// TIA Portal project "汽车系统" (V15.1)
// 汽车雨刷与车窗系统

(* hardware
DEVICE "S7-1200 station_1"  S7-1200 Station
   slot 0: "Rack_0"  S7-1200 Rack  Rack  V1.0
   slot 1: "plc左"  CPU 1214C DC/DC/DC  6ES7 214-1AG40-0XB0  V4.2
   slot 2: "DI 16/DQ 16x24VDC_1"  6ES7 223-1BL32-0XB0  V2.0
   slot 3: "AI 4x13BIT/AQ 2x14BIT_1"  6ES7 234-4HE32-0XB0  V2.0
DEVICE "S7-1200 station_2"  S7-1200 Station
   slot 0: "Rack_0"  S7-1200 Rack  Rack  V1.0
   slot 1: "plc右"  CPU 1214C DC/DC/DC  6ES7 214-1AG40-0XB0  V4.2
   slot 2: "DI 16/DQ 16x24VDC_1"  6ES7 223-1BL32-0XB0  V2.0
   slot 3: "AI 4x13BIT/AQ 2x14BIT_1"  6ES7 234-4HE32-0XB0  V2.0
DEVICE "g120"  GSD.Device.PN
   slot 0: "机架"  Rack  V1.0
   slot 0: "g120"  SINAMICS G120 CU250S-2 PN Vector V4.7  6SL3 246-0BA22-1FAx  V4.70
      slot 0: "SINAMICS G120 CU250S-2 PN Vector V4.7"  SINAMICS G120 CU250S-2 PN Vector V4.7
      slot 1: "PN-IO"  PN-IO
         slot 1: "端口1"  Port 1
         slot 2: "端口2"  Port 2
      slot 1: "DO 矢量_1"  DO VECTOR
         slot 0: "模块访问点"  Module Access Point
   slot 2: "标准报文3_PZD5_9"  Standard telegram 3, PZD-5/9
DEVICE "v90"  GSD.Device.PN
   slot 0: "机架"  Rack  V1.0
   slot 0: "v90"  SINAMICS V90 PN V1.0  6SL3 210-5Fxxx-xxFx  V1.00
      slot 0: "SINAMICS V90 PN V1.0"  SINAMICS V90 PN V1.0
      slot 1: "PN-IO"  PN-IO
         slot 1: "端口1"  Port 1
         slot 2: "端口2"  Port 2
      slot 1: "驱动_1"  Drive
         slot 0: "模块访问点"  Module Access Point
         slot 1: "没有 PROFIsafe"  without PROFIsafe
   slot 2: "标准报文3_PZD5_9"  Standard telegram 3, PZD-5/9
DEVICE "HMI"  KTP700 Basic PN
   slot 0: "HMI"  KTP700 Basic PN  6AV2 123-2GB03-0AX0  15.1.0.0
   slot 1: "HMI_RT_1"  KTP700 Basic PN  6AV2 123-2GB03-0AX0  15.1.0.0
   slot 5: "HMI.IE_CP_1"  PROFINET Interface  15.0.1.0
      slot 1: "PROFINET Interface_1"  PROFINET Interface
         slot 1: "Port_1"  Port
*)

// ===== PLC "plc左"  CPU 1214C DC/DC/DC =====

VAR_GLOBAL   // PLC tag table "默认变量表"
   "Tag__639268081140296448" AT %I8.0 : Bool;
   "Tag__639268081140453381" AT %I8.1 : Bool;
   "Tag__639268081140484476" AT %I8.2 : Bool;
   "Tag__639268081140514566" AT %I8.3 : Bool;
   "Tag__639268081140554565" AT %I8.4 : Bool;
   "Tag__639268081140589602" AT %I8.5 : Bool;
   "Tag__639268081140634777" AT %I8.6 : Bool;
   "Tag__639268081140684765" AT %I8.7 : Bool;
   "Tag__639268081140724801" AT %I9.0 : Bool;
   "Tag__639268081140754790" AT %I9.1 : Bool;
   "Tag__639268081140789825" AT %I9.2 : Bool;
   "Tag__639268081140814951" AT %I9.3 : Bool;
   "Tag__639268081140834948" AT %I9.4 : Bool;
   "Tag__639268081140860990" AT %I9.5 : Bool;
   "Tag__639268081140890986" AT %I9.6 : Bool;
   "Tag__639268081140910987" AT %I9.7 : Bool;
   "Tag__639268081145756808" AT %Q8.0 : Bool;
   "Tag__639268081145787808" AT %Q8.1 : Bool;
   "Tag__639268081145815161" AT %Q8.2 : Bool;
   "Tag__639268081145835184" AT %Q8.3 : Bool;
   "Tag__639268081145856321" AT %Q8.4 : Bool;
   "Tag__639268081145886347" AT %Q8.5 : Bool;
   "Tag__639268081145901382" AT %Q8.6 : Bool;
   "Tag__639268081145931410" AT %Q8.7 : Bool;
   "Tag__639268081145951421" AT %Q9.0 : Bool;
   "Tag__639268081145971411" AT %Q9.1 : Bool;
   "Tag__639268081145991411" AT %Q9.2 : Bool;
   "Tag__639268081146013352" AT %Q9.3 : Bool;
   "Tag__639268081146043352" AT %Q9.4 : Bool;
   "Tag__639268081146063350" AT %Q9.5 : Bool;
   "Tag__639268081146073348" AT %Q9.6 : Bool;
   "Tag__639268081146103454" AT %Q9.7 : Bool;
   "Tag__639268084247338622" AT %QW8 : Word;
END_VAR

DATA_BLOCK "扫描计时实例"   // DB1
{ S7_Optimized_Access := 'TRUE' }
VERSION : 5.0
// 文件定位：左PLC/02_扫描计时实例.scl；TIA块名：“扫描计时实例”。
//  本块属于V3简明；与另两版执行代码和参数完全相同，差别仅为注释组织。
//  建议从左PLC/00_Main.scl开始，再回到本块阅读。
// stored: InstanceOfName 扫描计时
"扫描计时"
BEGIN
END_DATA_BLOCK

DATA_BLOCK "左侧参数"   // DB5
{ S7_Optimized_Access := 'TRUE' }
VERSION : 4.0
   VAR
      实机调试完成 : Bool := FALSE;   // 旧确认位保留，当前总控不以它作为运行许可条件。
      双机接收硬件标识 : Hw_Io := 276;   // 左PLC接收右状态使用的HW_IO标识，本工程276。
      双机发送硬件标识 : Hw_Io := 275;   // 左PLC发送命令使用的HW_IO标识，本工程275。
      使用手操盒 : Bool := false;   // 默认FALSE，忽略实体S01～S16，由有效PC/HMI请求产生逻辑钥匙；TRUE时恢复实体输入。
   END_VAR
BEGIN
END_DATA_BLOCK

DATA_BLOCK "汽车总控实例"   // DB6
{ S7_Optimized_Access := 'TRUE' }
VERSION : 5.0
// 文件定位：左PLC/11_汽车总控实例.scl；TIA块名：“汽车总控实例”。
//  本块属于V3简明；与另两版执行代码和参数完全相同，差别仅为注释组织。
//  建议从左PLC/00_Main.scl开始，再回到本块阅读。
// stored: InstanceOfName 汽车总控
"汽车总控"
BEGIN
END_DATA_BLOCK

DATA_BLOCK "上位机命令"   // DB100
{ S7_Optimized_Access := 'FALSE' }
VERSION : 4.0
   VAR
      字 : Array[0..31] of Word;
   END_VAR
BEGIN
END_DATA_BLOCK

DATA_BLOCK "上位机状态"   // DB101
{ S7_Optimized_Access := 'FALSE' }
VERSION : 4.0
   VAR
      字 : Array[0..63] of Word;
      雨刷实际角度 : Real;   // DBD128，HMI直接显示角度。
      车窗实际角度 : Real;   // DBD132，总长度136字节。
   END_VAR
BEGIN
END_DATA_BLOCK

DATA_BLOCK "面板命令"   // DB102
{ S7_Optimized_Access := 'FALSE' }
VERSION : 4.0
   VAR
      字 : Array[0..15] of Word;
   END_VAR
BEGIN
END_DATA_BLOCK

FUNCTION_BLOCK "汽车总控"   // FB1, SCL
{ S7_Optimized_Access := 'TRUE' }
VERSION : 5.0
// 文件定位：左PLC/10_汽车总控.scl；TIA块名：“汽车总控”。
//  本块属于V3简明；与另两版执行代码和参数完全相同，差别仅为注释组织。
//  建议从左PLC/00_Main.scl开始，再回到本块阅读。
   VAR_INPUT
      计时步数 : Int;
   END_VAR
   VAR
      上位机快照 : Array[0..31] of Word;
      上位机候选帧 : Array[0..31] of Word;
      面板上次值 : Array[0..15] of Word;
      手操开关 : Array[1..16] of Bool;
      开关上次值 : Array[1..16] of Bool;
      开关上升沿 : Array[1..16] of Bool;
      双机接收帧 : Array[0..15] of Word;
      双机发送帧 : Array[0..15] of Word;
      曾收到上位机 : Bool;
      曾收到面板 : Bool;
      曾收到右侧 : Bool;
      首次扫描 : Bool := TRUE;
      上位机心跳年龄 : Int := 30000;
      面板心跳年龄 : Int := 30000;
      右侧心跳年龄 : Int := 30000;
      上位机心跳 : Word;
      面板协调字 : Word;
      右侧心跳 : Word;
      上次模式票 : Word;
      上次一次票 : Word;
      上次复位票 : Word;
      命令确认序号 : Word;
      模式确认票 : Word;
      一次确认票 : Word;
      复位确认票 : Word;
      右侧复位票 : Word;
      本机心跳 : Word;
      状态序号 : Word;
      模式 : Int;
      档位 : Int;
      操作来源 : Int;
      一次保持计时 : Int;
      复位保持计时 : Int;
      一次等待启动 : Bool;
      一次执行中 : Bool;
      一次开始次数 : Word;
      复位拒绝次数 : Word;
      防夹全开锁定 : Bool;
      软件停止锁定 : Bool;
      等待按钮释放 : Bool;
      手操原始输入 : Word;
      手操有效输出 : Word;
      状态标志 : Word;
      提示标志 : Word;
      双机读结果 : Int;
      双机写结果 : Int;
      一次拒绝次数 : Word;
      雨量等级 : Int;
      上位机等待释放 : Bool := TRUE;
      面板等待释放 : Bool := TRUE;
      状态发布计时 : Int;
   END_VAR
   VAR_TEMP
      下标 : Int;
      模式开关数量 : Int;
      新选模式开关 : Int;
      暂存序号 : Word;
      帧有效 : Bool;
      新上位机命令 : Bool;
      上位机在线 : Bool;
      面板在线 : Bool;
      右侧在线 : Bool;
      上位机控制会话 : Bool;
      面板控制会话 : Bool;
      两轴启动完成 : Bool;
      雨刷就绪 : Bool;
      车窗就绪 : Bool;
      软件许可 : Bool;
      新一次请求 : Bool;
      新复位请求 : Bool;
      模式冲突 : Bool;
      升降冲突 : Bool;
      向上 : Bool;
      向下 : Bool;
      模拟手在位 : Bool;
      雨刷开关 : Bool;
      运行许可 : Bool;
      雨量有效 : Bool;
      模拟雨量 : Int;
      车窗开度 : Int;
      上位机向上 : Bool;
      上位机向下 : Bool;
      面板向上 : Bool;
      面板向下 : Bool;
   END_VAR
BEGIN
       // 职责：PLC左的业务协调器。接收PC/HMI/可选手操输入，判断输入是否新鲜、请求是否合法，再形成四个运动意图。
       // 本块不直接调用G120/V90驱动指令；最终雨刷与车窗动作由右PLC/10_右侧联动.scl转入两个轴FB。

       // 【输入所有权】参数决定采用实体S01～S16还是软件会话。无手操盒分支把实体输入全部忽略，S13逻辑允许。
       IF "左侧参数".使用手操盒 THEN
           #手操开关[1] := "Tag__639268081140296448";
           #手操开关[2] := "Tag__639268081140453381";
           #手操开关[3] := "Tag__639268081140484476";
           #手操开关[4] := "Tag__639268081140514566";
           #手操开关[5] := "Tag__639268081140554565";
           #手操开关[6] := "Tag__639268081140589602";
           #手操开关[7] := "Tag__639268081140634777";
           #手操开关[8] := "Tag__639268081140684765";
           #手操开关[9] := "Tag__639268081140724801";
           #手操开关[10] := "Tag__639268081140754790";
           #手操开关[11] := "Tag__639268081140789825";
           #手操开关[12] := "Tag__639268081140814951";
           #手操开关[13] := "Tag__639268081140834948";
           #手操开关[14] := "Tag__639268081140860990";
           #手操开关[15] := "Tag__639268081140890986";
           #手操开关[16] := "Tag__639268081140910987";
       ELSE

           FOR #下标 := 1 TO 16 DO
               #手操开关[#下标] := FALSE;
           END_FOR;
           #手操开关[13] := TRUE;
       END_IF;
       #手操原始输入 := 0;
       FOR #下标 := 1 TO 16 DO
           #开关上升沿[#下标] := #手操开关[#下标] AND NOT #开关上次值[#下标] AND NOT #首次扫描;
           #开关上次值[#下标] := #手操开关[#下标];
           IF #手操开关[#下标] THEN
               #手操原始输入 := #手操原始输入 OR SHL(IN := W#16#0001, N := INT_TO_UINT(#下标 - 1));
           END_IF;
       END_FOR;
       #首次扫描 := FALSE;
       #软件许可 := NOT #手操开关[11];
       #新一次请求 := FALSE;
       #新复位请求 := FALSE;
       #上位机心跳年龄 := "计时更新"(当前 := #上位机心跳年龄, 步数 := #计时步数, 上限 := 30000);
       #面板心跳年龄 := "计时更新"(当前 := #面板心跳年龄, 步数 := #计时步数, 上限 := 30000);
       #右侧心跳年龄 := "计时更新"(当前 := #右侧心跳年龄, 步数 := #计时步数, 上限 := 30000);
       #一次保持计时 := "计时更新"(当前 := #一次保持计时, 步数 := - #计时步数, 上限 := 100);
       #复位保持计时 := "计时更新"(当前 := #复位保持计时, 步数 := - #计时步数, 上限 := 20);

       // 【DB100顺序锁】先读头序号→复制32字→检查头尾/重新读头。写入中的奇数帧或复制中变化的帧都不消费。
       #暂存序号 := "上位机命令".字[2];
       FOR #下标 := 0 TO 31 DO
           #上位机候选帧[#下标] := "上位机命令".字[#下标];
       END_FOR;
       #帧有效 := (#上位机候选帧[0] = W#16#CA71) AND (#上位机候选帧[1] = W#16#0400)
       AND (#暂存序号 = #上位机候选帧[2]) AND (#暂存序号 = #上位机候选帧[31])
       AND (#暂存序号 = "上位机命令".字[2]) AND (#暂存序号 <> 0)
       AND ((#暂存序号 AND W#16#0001) = 0) AND (#上位机候选帧[4] <= 4)
       AND (#上位机候选帧[5] <= 1000) AND ((#上位机候选帧[6] AND W#16#FFC0) = 0);
       FOR #下标 := 10 TO 30 DO
           IF #上位机候选帧[#下标] <> 0 THEN
               #帧有效 := FALSE;
           END_IF;
       END_FOR;
       #新上位机命令 := FALSE;
       // 【新帧与新事件】心跳变化才刷新年龄。首次/重连时只保存当前票号基线，下一份持续在线的新票才产生事件。
       IF #帧有效 AND ((NOT #曾收到上位机) OR (#上位机候选帧[3] <> #上位机心跳)) THEN
           #新上位机命令 := #曾收到上位机 AND (#上位机心跳年龄 < 60);
           IF NOT #新上位机命令 THEN
               #上次模式票 := #上位机候选帧[9];
               #上次一次票 := #上位机候选帧[7];
               #上次复位票 := #上位机候选帧[8];
           END_IF;
           FOR #下标 := 0 TO 31 DO
               #上位机快照[#下标] := #上位机候选帧[#下标];
           END_FOR;
           #曾收到上位机 := TRUE;
           #上位机心跳年龄 := 0;
           #上位机心跳 := #上位机候选帧[3];
           #命令确认序号 := #暂存序号;
       END_IF;

       #上位机在线 := #曾收到上位机 AND (#上位机心跳年龄 < 60);
       #上位机控制会话 := #上位机在线 AND #手操开关[13] AND #上位机快照[6].%X4;

       // 【HMI独立入口】DB102字0～4为模式翻转票，5一次，6/7升降保持，8防夹，9复位，10停止。
       IF "面板命令".字[12] <> #面板协调字 THEN
           IF NOT #曾收到面板 OR (#面板心跳年龄 >= 250) THEN
               FOR #下标 := 0 TO 15 DO
                   #面板上次值[#下标] := "面板命令".字[#下标];
               END_FOR;
           END_IF;
           #面板协调字 := "面板命令".字[12];
           #面板心跳年龄 := 0;
           #曾收到面板 := TRUE;
       END_IF;
       #面板在线 := #曾收到面板 AND (#面板心跳年龄 < 250);
       #面板控制会话 := #面板在线 AND #手操开关[13] AND "面板命令".字[11].%X0;
       IF NOT "左侧参数".使用手操盒 THEN

           #手操开关[1] := #上位机控制会话 OR #面板控制会话;

           #手操原始输入.%X0 := #手操开关[1];
           #手操原始输入.%X12 := TRUE;
       END_IF;

       // 【读取右侧】先校验DPRD_DAT返回码与D401/0400，再检查首尾心跳和开度范围。
       #双机读结果 := -1;
       IF "左侧参数".双机接收硬件标识 <> 0 THEN
           #双机读结果 := DPRD_DAT(LADDR := "左侧参数".双机接收硬件标识, RECORD => #双机接收帧);
       END_IF;
       #帧有效 := (#双机读结果 = 0) AND (#双机接收帧[0] = W#16#D401) AND (#双机接收帧[1] = W#16#0400)
       AND (#双机接收帧[2] = #双机接收帧[15]) AND ((#双机接收帧[4] <= 100) OR (#双机接收帧[4] = 255));

       IF (#双机接收帧[10] AND W#16#FF00) <> 0 THEN
           #帧有效 := FALSE;
       END_IF;
       IF #帧有效 AND ((NOT #曾收到右侧) OR (#双机接收帧[2] <> #右侧心跳)) THEN
           #曾收到右侧 := TRUE;
           #右侧心跳年龄 := 0;
           #右侧心跳 := #双机接收帧[2];
       END_IF;
       #右侧在线 := #曾收到右侧 AND (#右侧心跳年龄 < 30) AND #帧有效;
       #车窗开度 := 255;
       IF #右侧在线 THEN
           #车窗开度 := WORD_TO_INT(#双机接收帧[4]);
       END_IF;

       // 【独立就绪】雨刷接受质量bit0实测或bit7估算，再叠加雨刷启动完成；车窗要求bit1实际反馈及车窗启动完成。
       #雨刷就绪 := #右侧在线 AND (#双机接收帧[10].%X0 OR #双机接收帧[10].%X7) AND #双机接收帧[10].%X4;
       #车窗就绪 := #右侧在线 AND #双机接收帧[10].%X1 AND #双机接收帧[10].%X5;
       #两轴启动完成 := #雨刷就绪 AND #车窗就绪;

       // 【事件票据】票号变化表示一次新的用户意图。模式票消费后回显；一次和复位还各有接受条件和拒绝计数。
       IF #新上位机命令 THEN
           IF #上位机快照[9] <> #上次模式票 THEN
               IF #上位机控制会话 THEN
                   #模式 := WORD_TO_INT(#上位机快照[4]);
                   #操作来源 := 2;
               END_IF;
               #模式确认票 := #上位机快照[9];
           END_IF;
           IF #上位机快照[7] <> #上次一次票 THEN
               #新一次请求 := #上位机控制会话;
               #一次确认票 := #上位机快照[7];
           END_IF;
           IF #上位机快照[8] <> #上次复位票 THEN
               #新复位请求 := #上位机在线 AND #手操开关[13];
               #复位确认票 := #上位机快照[8];
           END_IF;
           #上次模式票 := #上位机快照[9];
           #上次一次票 := #上位机快照[7];
           #上次复位票 := #上位机快照[8];
       END_IF;
       IF (#操作来源 = 2) AND NOT #上位机控制会话 THEN
           #模式 := 0;
       END_IF;
       IF (#操作来源 = 3) AND NOT #面板控制会话 THEN
           #模式 := 0;
       END_IF;

       FOR #下标 := 0 TO 4 DO
           IF "面板命令".字[#下标] <> #面板上次值[#下标] THEN
               IF #面板控制会话 THEN
                   #模式 := #下标;
                   #操作来源 := 3;
               END_IF;
           END_IF;
       END_FOR;
       IF ("面板命令".字[5] <> #面板上次值[5]) AND #面板控制会话 THEN
           #新一次请求 := TRUE;
       END_IF;
       IF ("面板命令".字[9] <> #面板上次值[9]) AND #面板在线 AND #手操开关[13] THEN
           #新复位请求 := TRUE;
       END_IF;
       IF ("面板命令".字[10] <> #面板上次值[10]) AND #面板在线 THEN
           #软件停止锁定 := TRUE;
       END_IF;
       FOR #下标 := 0 TO 15 DO
           #面板上次值[#下标] := "面板命令".字[#下标];
       END_FOR;

       #模式开关数量 := 0;
       #新选模式开关 := 0;
       FOR #下标 := 2 TO 6 DO
           IF #手操开关[#下标] THEN
               #模式开关数量 := #模式开关数量 + 1;
           END_IF;
           IF #开关上升沿[#下标] THEN
               #新选模式开关 := #下标;
           END_IF;
       END_FOR;
       #模式冲突 := #模式开关数量 > 1;
       IF #新选模式开关 > 0 THEN
           #模式 := #新选模式开关 - 2;
           #操作来源 := 1;
       END_IF;
       IF #模式冲突 THEN
           #模式 := 0;
           #操作来源 := 1;
       END_IF;
       IF #开关上升沿[7] THEN
           #新一次请求 := TRUE;
       END_IF;
       IF #开关上升沿[10] THEN
           #新复位请求 := TRUE;
       END_IF;
       IF #手操开关[11] OR (#上位机在线 AND #上位机快照[6].%X3) THEN
           #软件停止锁定 := TRUE;
       END_IF;

       // 【自动档迟滞】只有雨量有效时参与自动选档。进入阈值50/350/700，退出阈值20/300/650。
       #雨量有效 := #上位机在线 AND #上位机快照[6].%X5;
       #模拟雨量 := 0;
       IF #雨量有效 THEN
           #模拟雨量 := WORD_TO_INT(#上位机快照[5]);
       END_IF;

       IF NOT #雨量有效 THEN
           #雨量等级 := 0;
       ELSE
           CASE #雨量等级 OF
               0:
                   IF #模拟雨量 >= 50 THEN
                       #雨量等级 := 1;
                   END_IF;
               1:
                   IF #模拟雨量 < 20 THEN
                       #雨量等级 := 0;
                   ELSIF #模拟雨量 >= 350 THEN
                       #雨量等级 := 2;
                   END_IF;
               2:
                   IF #模拟雨量 < 300 THEN
                       #雨量等级 := 1;
                   ELSIF #模拟雨量 >= 700 THEN
                       #雨量等级 := 3;
                   END_IF;
               3:
                   IF #模拟雨量 < 650 THEN
                       #雨量等级 := 2;
                   END_IF;
               ELSE
                   #雨量等级 := 0;
           END_CASE;
       END_IF;
       #档位 := 0;
       CASE #模式 OF
           1:
               #档位 := #雨量等级;
           2:
               #档位 := 1;
           3:
               #档位 := 2;
           4:
               #档位 := 3;
       END_CASE;

       // 【重新操作】会话重新建立后，先观察升降均释放，再允许新的保持命令。PC与HMI各有自己的释放记忆。
       IF NOT #上位机控制会话 THEN
           #上位机等待释放 := TRUE;
       ELSIF NOT #上位机快照[6].%X0 AND NOT #上位机快照[6].%X1 THEN
           #上位机等待释放 := FALSE;
       END_IF;
       IF NOT #面板控制会话 THEN
           #面板等待释放 := TRUE;
       ELSIF NOT "面板命令".字[6].%X0 AND NOT "面板命令".字[7].%X0 THEN
           #面板等待释放 := FALSE;
       END_IF;
       #上位机向上 := #上位机控制会话 AND NOT #上位机等待释放 AND #上位机快照[6].%X0;
       #上位机向下 := #上位机控制会话 AND NOT #上位机等待释放 AND #上位机快照[6].%X1;

       #面板向上 := #面板控制会话 AND NOT #面板等待释放 AND "面板命令".字[6].%X0;
       #面板向下 := #面板控制会话 AND NOT #面板等待释放 AND "面板命令".字[7].%X0;
       #向上 := #手操开关[8] OR #上位机向上 OR #面板向上;
       #向下 := #手操开关[9] OR #上位机向下 OR #面板向下;

       // 【防夹事件变任务】PC/HMI脉冲触发后锁定全开。即使UI脉冲和冷却按钮已经结束，PLC继续要求开窗。
       #模拟手在位 := #手操开关[12] OR (#上位机在线 AND #手操开关[13] AND #上位机快照[6].%X2)
       OR (#面板在线 AND #手操开关[13] AND "面板命令".字[8].%X0);
       IF #模拟手在位 THEN
           #防夹全开锁定 := TRUE;
           #等待按钮释放 := TRUE;
       END_IF;
       #升降冲突 := #向上 AND #向下 AND NOT #防夹全开锁定;
       IF #升降冲突 THEN
           #等待按钮释放 := TRUE;
       END_IF;
       IF NOT #向上 AND NOT #向下 AND NOT #模拟手在位 THEN
           #等待按钮释放 := FALSE;
       END_IF;
       IF #防夹全开锁定 AND (#车窗开度 = 100) AND NOT #模拟手在位 THEN
           #防夹全开锁定 := FALSE;
           #等待按钮释放 := TRUE;
       END_IF;

       // 【复位条件逐项看】逻辑钥匙关闭、上下释放、防夹释放、实体停止释放、软件许可成立且PC停止位清除。
       IF #新复位请求 THEN
           IF NOT #手操开关[1] AND NOT #向上 AND NOT #向下 AND NOT #模拟手在位
               AND NOT #手操开关[11] AND #软件许可
               AND NOT (#上位机在线 AND #上位机快照[6].%X3) THEN
               #软件停止锁定 := FALSE;
               #模式 := 0;
               #档位 := 0;
               #一次保持计时 := 0;
               #一次等待启动 := FALSE;
               #一次执行中 := FALSE;
               #右侧复位票 := "字计数递增"(原值 := #右侧复位票);
               #复位保持计时 := 20;
           ELSE
               #复位拒绝次数 := "字计数递增"(原值 := #复位拒绝次数);
           END_IF;
       END_IF;

       // 【总运行许可】逻辑钥匙与软件许可有效、软件停止锁定已解除即可形成许可；不把两轴就绪塞进这个总条件。
       #运行许可 := #手操开关[1] AND #软件许可 AND NOT #软件停止锁定;
       IF NOT #运行许可 THEN
           #等待按钮释放 := TRUE;
       END_IF;

       // 【一次是闭环握手】只在运行许可、雨刷单轴就绪、右侧状态10且没有正在执行的一次任务时接受。
       IF #新一次请求 THEN
           IF #运行许可 AND #雨刷就绪 AND (#双机接收帧[6] = 10)
               AND NOT #一次等待启动 AND NOT #一次执行中 THEN
               #一次等待启动 := TRUE;
               #一次保持计时 := 100;
               #一次开始次数 := #双机接收帧[5];
               #模式 := 0;
           ELSE
               #一次拒绝次数 := "字计数递增"(原值 := #一次拒绝次数);
           END_IF;
       END_IF;
       // 【等右侧确认】看到运动状态就改为一次执行中，并撤销继续启动意图；右PLC仍会完成已锁定的整轮。
       IF #一次等待启动 THEN
           IF #右侧在线 AND ((#双机接收帧[6] = 20) OR (#双机接收帧[6] = 21)
               OR (#双机接收帧[6] = 30) OR (#双机接收帧[6] = 31)) THEN
               #一次等待启动 := FALSE;
               #一次执行中 := TRUE;
               #一次保持计时 := 0;
           ELSIF #一次保持计时 = 0 THEN
               #一次等待启动 := FALSE;
               #一次拒绝次数 := "字计数递增"(原值 := #一次拒绝次数);
           END_IF;
       END_IF;
       IF #一次执行中 AND #右侧在线 AND (#双机接收帧[5] <> #一次开始次数) THEN
           #一次执行中 := FALSE;
       END_IF;

       // 【一次固定中档】档位2意味着正向10 s、反向10 s名义保持时间。开始后清继续启动开关，等待完成次数变化。
       IF #一次等待启动 OR #一次执行中 THEN
           #档位 := 2;
       END_IF;
       #雨刷开关 := (#档位 > 0) AND #运行许可 AND #雨刷就绪;
       IF #一次执行中 THEN
           #雨刷开关 := FALSE;
       END_IF;
       IF #等待按钮释放 OR NOT #车窗就绪 THEN
           #向上 := FALSE;
           #向下 := FALSE;
       END_IF;

       IF #防夹全开锁定 THEN
           #向上 := FALSE;
           #向下 := TRUE;
       END_IF;
       IF NOT #运行许可 OR NOT #右侧在线 THEN
           #向上 := FALSE;
           #向下 := FALSE;
           #雨刷开关 := FALSE;
           #一次保持计时 := 0;
           #一次等待启动 := FALSE;
           #一次执行中 := FALSE;
       END_IF;
       IF #复位保持计时 > 0 THEN
           #雨刷开关 := FALSE;
           #向上 := FALSE;
           #向下 := FALSE;
       END_IF;

       // 【C401发送映射】先清空16字，写魔数/版本/心跳；字3.bit0许可、bit1停止，字4复位票。
       #本机心跳 := "字计数递增"(原值 := #本机心跳);
       FOR #下标 := 0 TO 15 DO
           #双机发送帧[#下标] := 0;
       END_FOR;
       #双机发送帧[0] := W#16#C401;
       #双机发送帧[1] := W#16#0400;
       #双机发送帧[2] := #本机心跳;
       #双机发送帧[3].%X0 := #运行许可;
       #双机发送帧[3].%X1 := #软件停止锁定 OR NOT #软件许可;
       #双机发送帧[4] := #右侧复位票;
       #双机发送帧[5] := BOOL_TO_WORD(#雨刷开关);
       #双机发送帧[6] := INT_TO_WORD(#档位);
       #双机发送帧[7] := BOOL_TO_WORD(#向上);
       #双机发送帧[8] := BOOL_TO_WORD(#向下);
       #双机发送帧[15] := #本机心跳;
       #双机写结果 := -1;
       IF "左侧参数".双机发送硬件标识 <> 0 THEN
           #双机写结果 := DPWR_DAT(LADDR := "左侧参数".双机发送硬件标识, RECORD := #双机发送帧);
       END_IF;

       // 【指示输出】按最终仲裁结果填指示字，不是根据界面按钮颜色推断状态。
       #手操有效输出 := 0;
       #手操有效输出.%X0 := #运行许可;
       #手操有效输出.%X1 := #模式 = 0;
       #手操有效输出.%X2 := #模式 = 1;
       #手操有效输出.%X3 := #模式 = 2;
       #手操有效输出.%X4 := #模式 = 3;
       #手操有效输出.%X5 := #模式 = 4;
       #手操有效输出.%X6 := #一次等待启动 OR #一次执行中;
       #手操有效输出.%X7 := #向上;
       #手操有效输出.%X8 := #向下;
       #手操有效输出.%X9 := #车窗开度 = 0;
       #手操有效输出.%X10 := #车窗开度 = 100;
       #手操有效输出.%X11 := #防夹全开锁定;
       #手操有效输出.%X12 := #手操开关[13];
       #手操有效输出.%X13 := #右侧在线;
       #手操有效输出.%X14 := FALSE;
       #手操有效输出.%X15 := FALSE;
       "Tag__639268081145756808" := #手操有效输出.%X0;
       "Tag__639268081145787808" := #手操有效输出.%X1;
       "Tag__639268081145815161" := #手操有效输出.%X2;
       "Tag__639268081145835184" := #手操有效输出.%X3;
       "Tag__639268081145856321" := #手操有效输出.%X4;
       "Tag__639268081145886347" := #手操有效输出.%X5;
       "Tag__639268081145901382" := #手操有效输出.%X6;
       "Tag__639268081145931410" := #手操有效输出.%X7;
       "Tag__639268081145951421" := #手操有效输出.%X8;
       "Tag__639268081145971411" := #手操有效输出.%X9;
       "Tag__639268081145991411" := #手操有效输出.%X10;
       "Tag__639268081146013352" := #手操有效输出.%X11;
       "Tag__639268081146043352" := #手操有效输出.%X12;
       "Tag__639268081146063350" := #手操有效输出.%X13;

       "Tag__639268081146073348" := FALSE;
       "Tag__639268081146103454" := FALSE;
       #状态标志 := 0;
       #状态标志.%X0 := #手操开关[1];
       #状态标志.%X1 := #软件许可;
       #状态标志.%X2 := #上位机在线;
       #状态标志.%X3 := #右侧在线;
       #状态标志.%X4 := #上位机控制会话;
       #状态标志.%X5 := #雨刷开关;
       #状态标志.%X6 := #两轴启动完成;
       #状态标志.%X7 := #向上;
       #状态标志.%X8 := #向下;
       #状态标志.%X9 := #防夹全开锁定;
       #状态标志.%X10 := #模拟手在位;
       #状态标志.%X11 := #车窗开度 = 100;
       #状态标志.%X12 := #车窗开度 = 0;
       #状态标志.%X13 := #车窗开度 <= 100;
       #状态标志.%X14 := #运行许可;
       #状态标志.%X15 := #软件停止锁定;
       #提示标志 := 0;
       #提示标志.%X0 := NOT #雨量有效;
       #提示标志.%X1 := #模式冲突;
       #提示标志.%X2 := #升降冲突;
       #提示标志.%X3 := NOT #面板在线;
       #提示标志.%X4 := NOT #右侧在线;
       #提示标志.%X5 := NOT #两轴启动完成;
       #提示标志.%X6 := NOT #上位机在线;
       #提示标志.%X7 := #等待按钮释放 OR (#上位机控制会话 AND #上位机等待释放)
       OR (#面板控制会话 AND #面板等待释放);

       #状态发布计时 := "计时更新"(当前 := #状态发布计时, 步数 := #计时步数, 上限 := 10);

       // 【DB101发布顺序锁】每100 ms先置奇数头序号，写状态数据，最后写同一偶数尾序号与头序号。
       IF #状态发布计时 >= 10 THEN
           #状态发布计时 := 0;
           IF #状态序号 >= W#16#FFFE THEN
               #状态序号 := W#16#0002;
           ELSE
               #状态序号 := UINT_TO_WORD(WORD_TO_UINT(#状态序号) + UINT#2);
           END_IF;
           "上位机状态".字[2] := #状态序号 OR W#16#0001;
           "上位机状态".字[0] := W#16#CA72;
           "上位机状态".字[1] := W#16#0400;
           "上位机状态".字[3] := #本机心跳;
           "上位机状态".字[4] := #命令确认序号;
           "上位机状态".字[5] := #一次确认票;
           "上位机状态".字[6] := #复位确认票;
           "上位机状态".字[7] := INT_TO_WORD(#模式);
           "上位机状态".字[8] := INT_TO_WORD(#档位);
           "上位机状态".字[9] := INT_TO_WORD(#操作来源);
           "上位机状态".字[10] := #手操原始输入;
           "上位机状态".字[11] := INT_TO_WORD(#模拟雨量);
           "上位机状态".字[12] := #状态标志;
           "上位机状态".字[13] := #提示标志;
           "上位机状态".字[14] := #双机接收帧[3];
           "上位机状态".字[15] := #手操有效输出;
           "上位机状态".字[16] := INT_TO_WORD(#车窗开度);
           "上位机状态".字[17] := INT_TO_WORD(#一次保持计时);
           "上位机状态".字[18] := #一次拒绝次数;
           "上位机状态".字[19] := 0;
           "上位机状态".字[19].%X0 := #面板控制会话;
           "上位机状态".字[19].%X1 := #面板控制会话 AND #运行许可 AND #雨刷就绪 AND (#双机接收帧[6] = 10)
           AND NOT #一次等待启动 AND NOT #一次执行中;
           "上位机状态".字[19].%X2 := #面板控制会话 AND #运行许可 AND #车窗就绪 AND NOT #防夹全开锁定;
           "上位机状态".字[20] := #右侧心跳;
           "上位机状态".字[21] := #面板协调字;
           "上位机状态".字[22] := INT_TO_WORD(#上位机心跳年龄);
           "上位机状态".字[23] := INT_TO_WORD(#右侧心跳年龄);
           "上位机状态".字[24] := INT_TO_WORD(#面板心跳年龄);
           "上位机状态".字[25] := INT_TO_WORD(#双机写结果);
           "上位机状态".字[26] := INT_TO_WORD(#双机读结果);
           "上位机状态".字[27] := #模式确认票;
           "上位机状态".字[28] := "面板命令".字[13];
           FOR #下标 := 29 TO 62 DO
               "上位机状态".字[#下标] := 0;
           END_FOR;
           IF #右侧在线 THEN
               "上位机状态".字[29] := #双机接收帧[8];
               "上位机状态".字[30] := #双机接收帧[9];
               "上位机状态".字[31] := #双机接收帧[10];
               "上位机状态".字[32] := #双机接收帧[5];
               "上位机状态".字[33] := #双机接收帧[6];
               "上位机状态".字[34] := #双机接收帧[7];
               "上位机状态".字[35] := #双机接收帧[11];
               "上位机状态".字[36] := #双机接收帧[12];
               "上位机状态".字[37] := #双机接收帧[13];
               "上位机状态".字[38] := #双机接收帧[14];
           END_IF;
           "上位机状态".字[39].%X0 := #一次等待启动;
           "上位机状态".字[39].%X1 := #一次执行中;
           "上位机状态".字[39].%X2 := #雨刷就绪;
           "上位机状态".字[39].%X3 := #车窗就绪;
           "上位机状态".字[40] := #复位拒绝次数;
           "上位机状态".雨刷实际角度 := INT_TO_REAL(WORD_TO_INT("上位机状态".字[29])) / 100.0;
           "上位机状态".车窗实际角度 := INT_TO_REAL(WORD_TO_INT("上位机状态".字[30])) / 100.0;
           "上位机状态".字[63] := #状态序号;
           "上位机状态".字[2] := #状态序号;
       END_IF;
END_FUNCTION_BLOCK

FUNCTION_BLOCK "扫描计时"   // FB2, SCL
{ S7_Optimized_Access := 'TRUE' }
VERSION : 5.0
// 左PLC完整可导入SCL源码。阅读请从同目录的左PLC/00_Main.scl或本文件ORGANIZATION_BLOCK "Main"开始。
//  保留原始块顺序便于TIA依赖解析；下面的代码与其他两版本一致，只有中文说明与排版不同。
//  参数XML及现有TIA工程共同提供通信DB、工艺对象和原生MC实例；完整工程是下载使用入口。
//  文件定位：左PLC/01_扫描计时.scl；TIA块名：“扫描计时”。
//  本块属于V3简明；与另两版执行代码和参数完全相同，差别仅为注释组织。
//  建议从左PLC/00_Main.scl开始，再回到本块阅读。
   VAR_OUTPUT
      时间步数 : Int;
   END_VAR
   VAR
      时标 : LReal;
      不足十毫秒余量 : LReal;
      首次调用 : Bool := TRUE;
   END_VAR
   VAR_TEMP
      本周期秒 : LReal;
      完整步数 : DInt;
   END_VAR
BEGIN
       // 此FB把不固定的CPU扫描周期换算成统一10 ms步数。每个PLC都有自己的实例，不跨CPU共享时钟。
       // RUNTIME返回的是相邻调用之间的秒数，包含通信/中断消耗；首次只初始化，非正样本不累加。

       // 【计时来源】RUNTIME使用CPU时钟测相邻调用间隔，先读取再判断首样本；界面刷新快慢不会影响这里。
       #本周期秒 := RUNTIME(#时标);
       #时间步数 := 0;
       IF #首次调用 THEN
           #首次调用 := FALSE;
           #不足十毫秒余量 := 0.0;
       ELSIF #本周期秒 > 0.0 THEN
           #不足十毫秒余量 := #不足十毫秒余量 + #本周期秒;

           // 【饱和】300 s相当于30000个10 ms步，仍在INT正范围内，防止暂停后转换溢出。
           IF #不足十毫秒余量 >= 300.0 THEN
               #时间步数 := 30000;
               #不足十毫秒余量 := 0.0;
           ELSE
               // 【保留余量】只输出完整10 ms的部分，减去已输出时间，未满一格的余量下次继续用。
               #完整步数 := TRUNC_DINT(#不足十毫秒余量 / 0.01);
               #时间步数 := DINT_TO_INT(#完整步数);
               #不足十毫秒余量 := #不足十毫秒余量 - DINT_TO_LREAL(#完整步数) * 0.01;
           END_IF;
       END_IF;
END_FUNCTION_BLOCK

FUNCTION "字计数递增" : Word   // FC1, SCL
{ S7_Optimized_Access := 'TRUE' }
VERSION : 4.0
// 左侧完整用户源程序。导入后为命令/状态/面板/右屏DB手动指定100/101/102/103。
//  本源与右侧源分别导入对应CPU，不能在同一CPU重复生成同名函数。
   VAR_INPUT
      原值 : Word;
   END_VAR
BEGIN
       IF #原值 = W#16#FFFF THEN
           #字计数递增 := 0;
       ELSE
           #字计数递增 := UINT_TO_WORD(WORD_TO_UINT(#原值) + UINT#1);
       END_IF;
END_FUNCTION

FUNCTION "计时更新" : Int   // FC2, SCL
{ S7_Optimized_Access := 'TRUE' }
VERSION : 5.0
// 文件定位：左PLC/03_计时更新.scl；TIA块名：“计时更新”。
//  本块属于V3简明；与另两版执行代码和参数完全相同，差别仅为注释组织。
//  建议从左PLC/00_Main.scl开始，再回到本块阅读。
   VAR_INPUT
      当前 : Int;
      步数 : Int;
      上限 : Int;
   END_VAR
   VAR_TEMP
      新值 : DInt;
   END_VAR
BEGIN
       // 公共饱和计时FC，没有独立历史记忆：输入当前值、增量和上限，返回0～上限的INT。
       // 先把两个INT转DINT相加，再LIMIT，最后转回INT；加法不会先在INT中溢出。

       #新值 := INT_TO_DINT(#当前) + INT_TO_DINT(#步数);
       #计时更新 := DINT_TO_INT(LIMIT(MN := DINT#0, IN := #新值, MX := INT_TO_DINT(#上限)));
END_FUNCTION

ORGANIZATION_BLOCK "Main"   // OB1, SCL, ProgramCycle
{ S7_Optimized_Access := 'TRUE' }
VERSION : 5.0
// 文件定位：左PLC/00_Main.scl；TIA块名：“Main”。
//  本块属于V3简明；与另两版执行代码和参数完全相同，差别仅为注释组织。
   VAR_INPUT
      Initial_Call : Bool;   // Initial call of this OB
      Remanence : Bool;   // =True, if remanent data are available
   END_VAR
   VAR_TEMP
      时间步数 : Int;
   END_VAR
BEGIN
       // 阅读入口：本文件是左PLC的Main循环组织块。完整源在“左PLC_完整.scl”，分块入口在“左PLC/00_Main.scl”。
       // 调用顺序：Main → 扫描计时实例（FB扫描计时）→ 汽车总控实例（FB汽车总控）。
       // Main每扫描只获取一次时间，然后把同一时间步数传给本PLC的全部业务。时间步数为0也照常调用业务。
       // 第一跳：左PLC/01_扫描计时.scl；第二跳：左PLC/10_汽车总控.scl；第三跳：左PLC/03_计时更新.scl。
       // 实例DB说明分别在左PLC/02_扫描计时实例.scl、左PLC/11_汽车总控实例.scl。
       // 雨刷每半程小15 s、中10 s、大5 s；一次固定中档，正反向命令共20 s，换向仍等待原生停稳。
       // 车窗使用实际反馈的相对坐标，默认45度/秒，方向系数同时作用于指令与反馈。
       // 默认无手操盒。先释放动作与控制申请，复位得到接受后再申请运行。

       "扫描计时实例"(时间步数 => #时间步数);

       "汽车总控实例"(计时步数 := #时间步数);
END_ORGANIZATION_BLOCK

ORGANIZATION_BLOCK "启动初始化"   // OB100, SCL, Startup
{ S7_Optimized_Access := 'TRUE' }
VERSION : 5.0
// 文件定位：左PLC/90_启动初始化.scl；TIA块名：“启动初始化”。
//  本块属于V3简明；与另两版执行代码和参数完全相同，差别仅为注释组织。
//  建议从左PLC/00_Main.scl开始，再回到本块阅读。
   VAR_INPUT
      LostRetentive : Bool;   // True if retentive data are lost
      LostRTC : Bool;   // True if date and time are lost
   END_VAR
   VAR_TEMP
      下标 : Int;
   END_VAR
BEGIN
       // CPU启动时清通信基线、动作和时基，先锁停；复位接受后再申请控制。

       "左侧参数".实机调试完成 := FALSE;
       "汽车总控实例".首次扫描 := TRUE;
       "汽车总控实例".曾收到上位机 := FALSE;
       "汽车总控实例".曾收到面板 := FALSE;
       "汽车总控实例".曾收到右侧 := FALSE;
       "汽车总控实例".上位机心跳年龄 := 30000;
       "汽车总控实例".面板心跳年龄 := 30000;
       "汽车总控实例".右侧心跳年龄 := 30000;

       "汽车总控实例".软件停止锁定 := TRUE;
       "汽车总控实例".模式 := 0;
       "汽车总控实例".一次等待启动 := FALSE;
       "汽车总控实例".一次执行中 := FALSE;
       "汽车总控实例".一次保持计时 := 0;
       "汽车总控实例".复位保持计时 := 0;
       "汽车总控实例".防夹全开锁定 := FALSE;
       "汽车总控实例".等待按钮释放 := TRUE;
       "汽车总控实例".上位机等待释放 := TRUE;
       "汽车总控实例".面板等待释放 := TRUE;
       FOR #下标 := 0 TO 31 DO
           "上位机命令".字[#下标] := 0;
       END_FOR;
       FOR #下标 := 0 TO 63 DO
           "上位机状态".字[#下标] := 0;
       END_FOR;
       FOR #下标 := 0 TO 15 DO
           "面板命令".字[#下标] := 0;
       END_FOR;
       "上位机状态".字[16] := 255;
       "Tag__639268084247338622" := W#16#0000;

       "扫描计时实例".时标 := 0.0;
       "扫描计时实例".不足十毫秒余量 := 0.0;
       "扫描计时实例".首次调用 := TRUE;
       "扫描计时实例".时间步数 := 0;
END_ORGANIZATION_BLOCK

// ===== PLC "plc右"  CPU 1214C DC/DC/DC =====

VAR_GLOBAL   // PLC tag table "默认变量表"
   "雨刷轴_Drive_IN" AT %I256.0 : "PD_TEL3_IN";
   "雨刷轴_Drive_OUT" AT %Q256.0 : "PD_TEL3_OUT";
   "车窗轴_Drive_IN" AT %I288.0 : "PD_TEL3_IN";
   "车窗轴_Drive_OUT" AT %Q288.0 : "PD_TEL3_OUT";
END_VAR

DATA_BLOCK "右侧参数"   // DB12
{ S7_Optimized_Access := 'TRUE' }
VERSION : 4.0
   VAR
      实机调试完成 : Bool := FALSE;   // 兼容旧工程的确认位，当前业务不以它作为运行门槛。
      雨刷原生反馈核对完成 : Bool := FALSE;   // 旧确认位，当前雨刷速度模式不检查此位。
      车窗原生反馈核对完成 : Bool := FALSE;   // 旧确认位；当前车窗直接读取工艺对象的真实编码器状态。
      双机接收硬件标识 : Hw_Io := 292;   // DPRD_DAT使用的HW_IO标识，本工程292；不是I512地址值。
      双机发送硬件标识 : Hw_Io := 296;   // DPWR_DAT使用的HW_IO标识，本工程296；不是Q512地址值。
      维护模式 : Bool := FALSE;   // 旧参数保留兼容，不再用来同时暂停两个轴。
      雨刷原配绝对编码器 : Bool := FALSE;   // 旧MC_Home模式选择参数；本版雨刷不执行MC_Home，当前不用。
      车窗原配绝对编码器 : Bool := FALSE;   // 旧MC_Home模式选择参数；本版车窗使用相对定位，当前不用。
      雨刷标定申请 : Bool := FALSE;   // 旧参数保留；本版雨刷不需要标定，切换此位不会建立机械坐标。
      车窗标定申请 : Bool := FALSE;   // 使能、停稳、无定位/停止作业且升降释放时，FALSE→TRUE重新记录当前起点；完成后置FALSE。
      雨刷已知基准角度 : Real := -120.0;   // 旧标定参数保留，当前雨刷开环逻辑不使用。
      车窗已知基准角度 : Real := 0.0;   // 旧标定参数保留；本版记录当前起点为逻辑0°，不使用此值。
      雨刷低档速度 : Real := 60.0;   // 小档速度，单位度/秒，默认60；新周期开始时读取，范围至少5且不高于中档。
      雨刷中档速度 : Real := 120.0;   // 中档速度，单位度/秒，默认120；不得低于小档或高于大档。
      雨刷高档速度 : Real := 180.0;   // 大档速度，单位度/秒，默认180；不得超过雨刷轴最大速度180。
      雨刷回位速度 : Real := 5.0;   // 旧定位参数保留；本版正反转沿用同一周期速度，不使用单独回位速度。
      车窗运动速度 : Real := 45.0;   // 正常升降速度，单位度/秒，默认45，范围大于0且不超过60；180°理想行程4秒。
      车窗回位速度 : Real := 5.0;   // 仅兼容旧状态5/6，范围大于0且不超过30；正常运行使用车窗运动速度。
      到位允许误差 : Real := 0.5;   // 车窗目标与实际相对位置的允许误差，单位度，默认0.5；范围大于0且不超过1。
      停稳速度阈值 : Real := 0.5;   // 车窗判断停稳时允许的绝对实际速度，单位度/秒，默认0.5，还须原生StandStill为TRUE。
      车窗方向反转 : Bool := true;   // 默认TRUE。记录起点时锁定为方向系数-1，同时反转指令与反馈坐标；修改后需重记起点。
      雨刷开环时间系数 : Real := 1.0;   // 兼容基座的保留字段；本版本慢、中、快每个半程固定为15、10、5秒。
   END_VAR
BEGIN
END_DATA_BLOCK

DATA_BLOCK "右侧运行"   // DB13
{ S7_Optimized_Access := 'TRUE' }
VERSION : 4.0
   VAR
      网络有效 : Bool;
      联动许可 : Bool;
      软件停止 : Bool;
      复位请求 : Bool;
      雨刷开关 : Bool;
      雨刷档位 : Int;
      车窗向上 : Bool;
      车窗向下 : Bool;
   END_VAR
BEGIN
END_DATA_BLOCK

DATA_BLOCK "右侧状态"   // DB14
{ S7_Optimized_Access := 'TRUE' }
VERSION : 4.0
   VAR
      雨刷状态 : Int;
      车窗状态 : Int;
      雨刷实际角度 : Real;
      车窗实际角度 : Real;
      雨刷位置有效 : Bool;
      车窗位置有效 : Bool;
      雨刷启动完成 : Bool;
      车窗启动完成 : Bool;
      雨刷故障码 : Word;
      车窗故障码 : Word;
      雨刷完成次数 : Word;
      车窗开度 : USInt := 255;
   END_VAR
BEGIN
END_DATA_BLOCK

DATA_BLOCK "雨刮器实例"   // DB15
{ S7_Optimized_Access := 'TRUE' }
VERSION : 6.0
// 文件定位：右PLC/21_雨刮器实例.scl；TIA块名：“雨刮器实例”。
//  本块属于V3简明；与另两版执行代码和参数完全相同，差别仅为注释组织。
//  建议从右PLC/00_Main.scl开始，再回到本块阅读。
// stored: InstanceOfName 雨刮器
"雨刮器"
BEGIN
END_DATA_BLOCK

DATA_BLOCK "车窗实例"   // DB16
{ S7_Optimized_Access := 'TRUE' }
VERSION : 5.0
// 文件定位：右PLC/31_车窗实例.scl；TIA块名：“车窗实例”。
//  本块属于V3简明；与另两版执行代码和参数完全相同，差别仅为注释组织。
//  建议从右PLC/00_Main.scl开始，再回到本块阅读。
// stored: InstanceOfName 车窗
"车窗"
BEGIN
END_DATA_BLOCK

DATA_BLOCK "右侧联动实例"   // DB17
{ S7_Optimized_Access := 'TRUE' }
VERSION : 5.0
// 文件定位：右PLC/11_右侧联动实例.scl；TIA块名：“右侧联动实例”。
//  本块属于V3简明；与另两版执行代码和参数完全相同，差别仅为注释组织。
//  建议从右PLC/00_Main.scl开始，再回到本块阅读。
// stored: InstanceOfName 右侧联动
"右侧联动"
BEGIN
END_DATA_BLOCK

DATA_BLOCK "扫描计时实例"   // DB18
{ S7_Optimized_Access := 'TRUE' }
VERSION : 5.0
// 文件定位：右PLC/02_扫描计时实例.scl；TIA块名：“扫描计时实例”。
//  本块属于V3简明；与另两版执行代码和参数完全相同，差别仅为注释组织。
//  建议从右PLC/00_Main.scl开始，再回到本块阅读。
// stored: InstanceOfName 扫描计时
"扫描计时"
BEGIN
END_DATA_BLOCK

DATA_BLOCK "雨刷轴"   // DB1, Motion_DB
{ S7_Optimized_Access := 'TRUE' }
AUTHOR : SIMATIC
FAMILY : BasicMC
NAME : TO_PosAx
VERSION : 6.0
// stored: InstanceOfName TO_PositioningAxis
"TO_PositioningAxis"
BEGIN
   // Axis.Encoder.TelegramAddressOutCU = %Q256.0
   // Axis.Encoder.DoNameCU = g120.DO 矢量_1_编码器1
   // Axis.Encoder.TelegramAddressInCU = %I256.0
   // Axis.Drive.TelegramAddressOutCU = %Q256.0
   // Axis.Drive.TelegramType = 2
   // Axis.Drive.DoNameCU = g120.DO 矢量_1
   // Axis.Drive.TelegramAddressInCU = %I256.0
   // Axis.LengthUnit.LastDistance = 1005
   // Axis.Encoder.DbTypeCU = Classic
   // Axis.Drive.DbTypeCU = Classic
   // Axis.LengthUnitNormalized.Time = 1
   // Axis.LengthUnitNormalized.Distance = -2
   // Axis.Encoder.SelectedHscIndexCU = -1
END_DATA_BLOCK

DATA_BLOCK "车窗轴"   // DB2, Motion_DB
{ S7_Optimized_Access := 'TRUE' }
AUTHOR : SIMATIC
FAMILY : BasicMC
NAME : TO_PosAx
VERSION : 6.0
// stored: InstanceOfName TO_PositioningAxis
"TO_PositioningAxis"
BEGIN
   // Axis.Encoder.TelegramAddressOutCU = %Q288.0
   // Axis.Encoder.DoNameCU = v90.驱动_1_编码器1
   // Axis.Encoder.TelegramAddressInCU = %I288.0
   // Axis.Drive.TelegramAddressOutCU = %Q288.0
   // Axis.Drive.TelegramType = 2
   // Axis.Drive.DoNameCU = v90.驱动_1
   // Axis.Drive.TelegramAddressInCU = %I288.0
   // Axis.LengthUnit.LastDistance = 1005
   // Axis.Encoder.DbTypeCU = Classic
   // Axis.Drive.DbTypeCU = Classic
   // Axis.LengthUnitNormalized.Time = 1
   // Axis.LengthUnitNormalized.Distance = -2
   // Axis.Encoder.SelectedHscIndexCU = -1
END_DATA_BLOCK

FUNCTION_BLOCK "雨刮器"   // FB1, SCL
{ S7_Optimized_Access := 'TRUE' }
VERSION : 6.0
// 文件定位：右PLC/20_雨刮器.scl；TIA块名：“雨刮器”。
//  本块属于V3简明；与另两版执行代码和参数完全相同，差别仅为注释组织。
//  建议从右PLC/00_Main.scl开始，再回到本块阅读。
   VAR_INPUT
      开关 : Bool;
      档位 : Int;
      计时步数 : Int;
   END_VAR
   VAR
      状态 : Int;
      故障锁定 : Bool;
      故障码 : Word;
      启动完成 : Bool;
      完成次数 : Word;
      复位等待计时 : Int;
      行程计时 : Int;
      停稳计时 : Int;
      行程时限 : Int;
      定位速度 : Real := 60.0;
      估算角度 : Real := -120.0;
      估算有效 : Bool;
      相对基准有效 : Bool;
      相对原点 : Real;
      上次标定申请 : Bool;
      使能完成 : Bool;
      点动忙 : Bool;
      达到速度 : Bool;
      点动中断 : Bool;
      使能出错 : Bool;
      复位出错 : Bool;
      点动出错 : Bool;
      使能错误码 : Word;
      复位错误码 : Word;
      点动错误码 : Word;
   END_VAR
   VAR_TEMP
      基础许可 : Bool;
      请求使能 : Bool;
      正向 : Bool;
      反向 : Bool;
      原生停稳 : Bool;
      原生故障 : Bool;
      参数有效 : Bool;
   END_VAR
BEGIN
       // 职责：G120实验电机的非位置控制速度往返。调用链为Main→右侧联动→雨刮器实例→原生MC指令。
       // 原先定位控制发生跟随误差时，本实现改用MC_Power StartMode=0、MC_MoveJog PositionControlled=FALSE。

       // 【方向每扫描重算】上一扫描的正反转命令不自动续用；只有当前有效状态能重新置对应方向。
       #正向 := FALSE;
       #反向 := FALSE;
       #复位等待计时 := "计时更新"(当前 := #复位等待计时, 步数 := - #计时步数, 上限 := 30);
       #基础许可 := "右侧运行".网络有效 AND "右侧运行".联动许可 AND NOT "右侧运行".软件停止;
       #原生故障 := "雨刷轴".StatusBits.Error;
       #原生停稳 := "雨刷轴".StatusBits.Standstill AND NOT #点动忙;

       // 【复位不发运动】清业务锁存并回状态0，随后300 ms给MC_Reset处理；复位前上层已要求动作和许可释放。
       IF "右侧运行".复位请求 THEN
           #故障锁定 := FALSE;
           #故障码 := 0;
           #状态 := 0;
           #启动完成 := FALSE;
           #复位等待计时 := 30;
       END_IF;

       // 【速度参数】低档至少5，中档不低于低档，高档不低于中档且最大180度/秒。
       #参数有效 := ("右侧参数".雨刷低档速度 >= 5.0)
       AND ("右侧参数".雨刷中档速度 >= "右侧参数".雨刷低档速度)
       AND ("右侧参数".雨刷高档速度 >= "右侧参数".雨刷中档速度)
       AND ("右侧参数".雨刷高档速度 <= 180.0);
       IF NOT #故障锁定 AND NOT #参数有效 THEN
           #故障锁定 := TRUE;
           #故障码 := W#16#F005;
       END_IF;
       IF NOT #故障锁定 AND ((#状态 = 21) OR (#状态 = 31)) AND (#行程时限 <= 0) THEN
           #故障锁定 := TRUE;
           #故障码 := W#16#F005;
       END_IF;
       IF NOT #故障锁定 AND #原生故障 AND #基础许可 AND (#复位等待计时 = 0) THEN
           #故障锁定 := TRUE;
           #故障码 := W#16#F001;
       END_IF;
       IF NOT #故障锁定 AND "雨刷轴".StatusBits.ControlPanelActive AND #基础许可 THEN
           #故障锁定 := TRUE;
           #故障码 := W#16#F007;
       END_IF;
       // 【使能条件】有效网络、联动许可、无停止、无本轴锁存故障且复位等待结束。使能完成不代表已经选档转动。
       #请求使能 := #基础许可 AND NOT #故障锁定 AND (#复位等待计时 = 0);
       IF NOT #请求使能 THEN
           #状态 := 0;
           #启动完成 := FALSE;
           #行程计时 := 0;
           #停稳计时 := 0;
       ELSIF #使能完成 THEN
           CASE #状态 OF

                   // 【状态0】等原生停稳和Power.Status，记录诊断参考位置，并把显示估算设为-120度，随后待命。
               0:
                   IF #原生停稳 THEN
                       #相对原点 := "雨刷轴".ActualPosition;
                       #相对基准有效 := TRUE;
                       #估算角度 := -120.0;
                       #估算有效 := TRUE;
                       #启动完成 := TRUE;
                       #状态 := 10;
                   END_IF;

                   // 【状态10】这里才采样新周期档位；周期中只使用已经保存的定位速度和行程时限。
               10:
                   IF #开关 AND (#档位 >= 1) AND (#档位 <= 3) THEN

                       // 【三档固定半程】小1500×10 ms、中1000×10 ms、大500×10 ms；每个方向的指令保持与UI刷新无关。
                       CASE #档位 OF
                           1:
                               #定位速度 := "右侧参数".雨刷低档速度;
                               #行程时限 := 1500;
                           2:
                               #定位速度 := "右侧参数".雨刷中档速度;
                               #行程时限 := 1000;
                           3:
                               #定位速度 := "右侧参数".雨刷高档速度;
                               #行程时限 := 500;
                       END_CASE;

                       #行程计时 := 0;
                       #状态 := 20;
                   END_IF;
                   // 【状态20→21】发出正向命令的起始扫描，把行程计时清零，然后在21持续保持。
               20:
                   #正向 := TRUE;
                   #行程计时 := 0;
                   #状态 := 21;

                   // 【状态21】以真实10 ms步数累计正向时间，包含实际驱动加速阶段；达到时限撤销正向并进入停稳等待。
               21:
                   #正向 := TRUE;
                   #行程计时 := "计时更新"(当前 := #行程计时, 步数 := #计时步数, 上限 := #行程时限);
                   #估算角度 := -120.0 + 240.0 * INT_TO_REAL(#行程计时) / INT_TO_REAL(#行程时限);
                   IF #行程计时 >= #行程时限 THEN
                       // 【方向每扫描重算】上一扫描的正反转命令不自动续用；只有当前有效状态能重新置对应方向。
                       #正向 := FALSE;
                       #停稳计时 := 0;
                       #估算角度 := 120.0;
                       #状态 := 22;
                   END_IF;

                   // 【状态22】等待StatusBits.StandStill且MoveJog不忙，才允许反向；等满10 s仍未停稳报F004。
               22:
                   #停稳计时 := "计时更新"(当前 := #停稳计时, 步数 := #计时步数, 上限 := 1000);
                   IF #原生停稳 THEN
                       #状态 := 30;
                   ELSIF #停稳计时 >= 1000 THEN
                       #故障锁定 := TRUE;
                       #故障码 := W#16#F004;
                   END_IF;
                   // 【状态30→31】正向已经确认停稳，才发反向并清本方向计时。
               30:
                   #反向 := TRUE;
                   #行程计时 := 0;
                   #状态 := 31;

                   // 【状态31】使用本轮同一速度和时限反转；显示角度按时间从120回到-120，不测量实际回到相同机械角度。
               31:
                   #反向 := TRUE;
                   #行程计时 := "计时更新"(当前 := #行程计时, 步数 := #计时步数, 上限 := #行程时限);
                   #估算角度 := 120.0 - 240.0 * INT_TO_REAL(#行程计时) / INT_TO_REAL(#行程时限);
                   IF #行程计时 >= #行程时限 THEN
                       #反向 := FALSE;
                       #停稳计时 := 0;
                       #估算角度 := -120.0;
                       #状态 := 32;
                   END_IF;

                   // 【状态32】反向停稳后才使完成次数递增；左PLC一次任务依据次数变化结束，而不是依据UI动画到终点。
               32:
                   #停稳计时 := "计时更新"(当前 := #停稳计时, 步数 := #计时步数, 上限 := 1000);
                   IF #原生停稳 THEN
                       #完成次数 := "字计数递增"(原值 := #完成次数);
                       #状态 := 10;
                   ELSIF #停稳计时 >= 1000 THEN
                       #故障锁定 := TRUE;
                       #故障码 := W#16#F004;
                   END_IF;
               ELSE
                   #状态 := 0;
           END_CASE;
       END_IF;
       IF #故障锁定 THEN
           #状态 := 90;
           #启动完成 := FALSE;
           #请求使能 := FALSE;
           #正向 := FALSE;
           #反向 := FALSE;
       END_IF;

       // 【原生速度模式】Power.StartMode=0，下面MoveJog.PositionControlled=FALSE。三个MC实例每扫描调用，Enable/方向由上面状态机给出。
       "雨刷使能"(Axis := "雨刷轴",
              Enable := #请求使能,
              StartMode := 0,
              StopMode := 0,
              Status => #使能完成,
              Error => #使能出错,
              ErrorID => #使能错误码);
       "雨刷复位"(Axis := "雨刷轴",
              Execute := "右侧运行".复位请求,
              Restart := FALSE,
              Error => #复位出错,
              ErrorID => #复位错误码);
       "雨刷速度点动"(Axis := "雨刷轴",
                JogForward := #正向,
                JogBackward := #反向,
                Velocity := #定位速度,
                PositionControlled := FALSE,
                InVelocity => #达到速度,
                Busy => #点动忙,
                CommandAborted => #点动中断,
                Error => #点动出错,
                ErrorID => #点动错误码);

       // 【保存故障来源】先发生的业务故障保留；原生MC错误返回原始ErrorID，F001只是工艺对象总故障入口。
       IF NOT #故障锁定 AND #复位出错 THEN
           #故障锁定 := TRUE;
           #故障码 := #复位错误码;
       END_IF;
       IF NOT #故障锁定 AND #使能出错 AND (#复位等待计时 = 0) THEN
           #故障锁定 := TRUE;
           #故障码 := #使能错误码;
       END_IF;
       IF NOT #故障锁定 AND #点动出错 AND (#复位等待计时 = 0) THEN
           #故障锁定 := TRUE;
           #故障码 := #点动错误码;
       END_IF;
       IF NOT #故障锁定 AND #点动中断 AND (#正向 OR #反向) AND #请求使能 THEN
           #故障锁定 := TRUE;
           #故障码 := W#16#F006;
       END_IF;
       "右侧状态".雨刷状态 := #状态;

       "右侧状态".雨刷实际角度 := "雨刷轴".ActualPosition - #相对原点 - 120.0;
       "右侧状态".雨刷位置有效 := ("雨刷轴".StatusSensor[1].State = 2) AND #相对基准有效;
       "右侧状态".雨刷启动完成 := #启动完成 AND NOT #故障锁定;
       "右侧状态".雨刷故障码 := #故障码;
       "右侧状态".雨刷完成次数 := #完成次数;
END_FUNCTION_BLOCK

FUNCTION_BLOCK "车窗"   // FB2, SCL
{ S7_Optimized_Access := 'TRUE' }
VERSION : 5.0
// 文件定位：右PLC/30_车窗.scl；TIA块名：“车窗”。
//  本块属于V3简明；与另两版执行代码和参数完全相同，差别仅为注释组织。
//  建议从右PLC/00_Main.scl开始，再回到本块阅读。
   VAR_INPUT
      向上 : Bool;
      向下 : Bool;
      计时步数 : Int;
   END_VAR
   VAR_OUTPUT
      位置 : USInt := 255;
   END_VAR
   VAR
      状态 : Int;
      故障锁定 : Bool;
      故障码 : Word;
      启动完成 : Bool;
      动作计时 : Int;
      停稳计时 : Int;
      复位等待计时 : Int;
      上次标定申请 : Bool;
      相对基准有效 : Bool;
      相对原点 : Real;
      相对距离 : Real;
      方向系数 : Real := -1.0;
      目标角度 : Real;
      定位速度 : Real := 5.0;
      使能完成 : Bool;
      定位完成 : Bool;
      定位忙 : Bool;
      定位中断 : Bool;
      停止完成 : Bool;
      停止忙 : Bool;
      标定完成 : Bool;
      标定忙 : Bool;
      使能出错 : Bool;
      定位出错 : Bool;
      停止出错 : Bool;
      复位出错 : Bool;
      标定出错 : Bool;
      使能错误码 : Word;
      定位错误码 : Word;
      停止错误码 : Word;
      复位错误码 : Word;
      标定错误码 : Word;
   END_VAR
   VAR_TEMP
      执行定位 : Bool;
      执行停止 : Bool;
      执行标定 : Bool;
      请求使能 : Bool;
      基础许可 : Bool;
      反馈有效 : Bool;
      已有基准 : Bool;
      原生故障 : Bool;
      原生停稳 : Bool;
      标定方式 : Int;
      速度 : Real;
      角度 : Real;
      原始角度 : Real;
      满足到位 : Bool;
      开度整数 : Int;
   END_VAR
BEGIN
       // 职责：V90车窗相对位置控制。上下请求来自左PLC仲裁，本块独立完成使能、记录起点、位移、停车和反馈。
       // 首次使能并停稳后读取ActualPosition为相对原点，逻辑角度=(原生位置-相对原点)×方向系数。

       #执行定位 := FALSE;
       #执行停止 := FALSE;
       #执行标定 := FALSE;
       #复位等待计时 := "计时更新"(当前 := #复位等待计时, 步数 := - #计时步数, 上限 := 30);

       // 【实际位置链】ActualPosition→减本次相对原点→乘锁定方向系数→逻辑角度，显示和运动用同一坐标定义。
       #原始角度 := "车窗轴".ActualPosition;
       #角度 := (#原始角度 - #相对原点) * #方向系数;
       #速度 := "车窗轴".ActualVelocity;
       #原生故障 := "车窗轴".StatusBits.Error;

       #反馈有效 := "车窗轴".StatusSensor[1].State = 2;
       IF NOT #反馈有效 THEN
           #相对基准有效 := FALSE;
       END_IF;
       #已有基准 := #相对基准有效;
       #原生停稳 := "车窗轴".StatusBits.Standstill
       AND (ABS(#速度) <= "右侧参数".停稳速度阈值);

       #基础许可 := "右侧运行".网络有效 AND "右侧运行".联动许可
       AND NOT "右侧运行".软件停止;

       // 【复位清业务状态】保留原生反馈读取，清故障/动作等待，再等待300 ms处理原生Reset。
       IF "右侧运行".复位请求 THEN
           #故障锁定 := FALSE;
           #故障码 := 0;
           #状态 := 0;
           #启动完成 := FALSE;
           #动作计时 := 0;
           #复位等待计时 := 30;
       END_IF;
       IF #原生故障 AND #基础许可 AND (#复位等待计时 = 0) THEN
           #故障锁定 := TRUE;
           #故障码 := W#16#F001;
       END_IF;
       IF (#启动完成 OR (#状态 = 6) OR (#状态 = 21) OR (#状态 = 31))
           AND NOT (#反馈有效 AND #已有基准) THEN
           #故障锁定 := TRUE;
           #故障码 := W#16#F002;
       END_IF;
       IF NOT (("右侧参数".到位允许误差 > 0.0) AND ("右侧参数".到位允许误差 <= 1.0)
           AND ("右侧参数".停稳速度阈值 > 0.0) AND ("右侧参数".停稳速度阈值 <= 1.0)) THEN
           #故障锁定 := TRUE;
           #故障码 := W#16#F005;
       END_IF;
       IF NOT (("右侧参数".车窗回位速度 > 0.0) AND ("右侧参数".车窗回位速度 <= 30.0)
           AND ("右侧参数".车窗运动速度 > 0.0) AND ("右侧参数".车窗运动速度 <= 60.0)) THEN
           #故障锁定 := TRUE;
           #故障码 := W#16#F005;
       END_IF;
       IF "车窗轴".StatusBits.ControlPanelActive AND #基础许可 THEN
           #故障锁定 := TRUE;
           #故障码 := W#16#F007;
       END_IF;
       #请求使能 := #基础许可 AND #反馈有效 AND NOT #故障锁定 AND (#复位等待计时 = 0);

       // 【记录任意起点】本轴使能、实际停稳、无定位/停止作业时记录；正常首次自动执行，重新标定须升降释放且申请有上升沿。
       IF #请求使能 AND #使能完成 AND #原生停稳 AND NOT #定位忙 AND NOT #停止忙
           AND ((NOT #相对基准有效)
           OR (NOT #向上 AND NOT #向下 AND "右侧参数".车窗标定申请 AND NOT #上次标定申请)) THEN

           IF "右侧参数".车窗方向反转 THEN
               #方向系数 := -1.0;
           ELSE
               #方向系数 := 1.0;
           END_IF;
           #相对原点 := #原始角度;
           #相对基准有效 := TRUE;
           #执行标定 := TRUE;
           #角度 := 0.0;
       END_IF;
       #已有基准 := #相对基准有效;
       #上次标定申请 := "右侧参数".车窗标定申请;
       IF NOT #请求使能 OR #执行标定 OR #标定忙 THEN
           #状态 := 0;
           #启动完成 := FALSE;
           #动作计时 := 0;
       ELSIF #使能完成 AND #已有基准 THEN
           // 【三个到位条件】Done说明相对定位指令完成，StandStill/实际速度确认已停，位置误差确认目标一致。
           #满足到位 := #定位完成 AND #原生停稳
           AND (ABS(#角度 - #目标角度) <= "右侧参数".到位允许误差);

           IF ((#状态 = 6) AND #向下)
               OR ((#状态 = 21) AND (NOT #向上 OR #向下))
               OR ((#状态 = 31) AND (NOT #向下 OR #向上)) THEN
               #启动完成 := TRUE;
               #状态 := 40;
           END_IF;

           // 【定位与停车状态】发令只在20/30计算一次相对距离，21/31保持等待；松手或换向先进入40/41停止。
           CASE #状态 OF
               0:
                   #启动完成 := TRUE;
                   #状态 := 10;
               5:
                   IF #向下 THEN
                       #启动完成 := TRUE;
                       #状态 := 30;
                   ELSE
                       #目标角度 := 0.0;
                       #定位速度 := "右侧参数".车窗回位速度;
                       #相对距离 := (#目标角度 - #角度) * #方向系数;
                       #执行定位 := TRUE;
                       #状态 := 6;
                   END_IF;
               6:
                   IF #满足到位 THEN
                       #启动完成 := TRUE;
                       #状态 := 10;
                   END_IF;
               10:
                   IF #向上 AND NOT #向下 AND (#角度 > "右侧参数".到位允许误差) THEN
                       #状态 := 20;
                   ELSIF #向下 AND NOT #向上 AND (#角度 < 180.0 - "右侧参数".到位允许误差) THEN
                       #状态 := 30;
                   END_IF;
                   // 【关窗发令】目标0度，距离=(0-当前逻辑角度)×方向系数，速度从车窗运动速度参数取。
               20:
                   IF #向上 AND NOT #向下 THEN
                       #目标角度 := 0.0;
                       #定位速度 := "右侧参数".车窗运动速度;
                       #相对距离 := (#目标角度 - #角度) * #方向系数;
                       #执行定位 := TRUE;
                       #状态 := 21;
                   ELSE
                       #状态 := 10;
                   END_IF;
               21:
                   IF #满足到位 THEN
                       #状态 := 10;
                   END_IF;
                   // 【开窗发令】目标180度，距离=(180-当前逻辑角度)×方向系数。
               30:
                   IF #向下 AND NOT #向上 THEN
                       #目标角度 := 180.0;
                       #定位速度 := "右侧参数".车窗运动速度;
                       #相对距离 := (#目标角度 - #角度) * #方向系数;
                       #执行定位 := TRUE;
                       #状态 := 31;
                   ELSE
                       #状态 := 10;
                   END_IF;
               31:
                   IF #满足到位 THEN
                       #状态 := 10;
                   END_IF;
               40:
                   #执行停止 := TRUE;
                   #状态 := 41;
               41:
                   IF #停止完成 AND #原生停稳 THEN
                       #状态 := 10;
                   END_IF;
               ELSE
                   #状态 := 0;
           END_CASE;
       END_IF;

       // 【Execute握手】在6/21/31等待态持续TRUE，让Done与稍后停稳能一起被消费；退出后释放，下一段再产生新上升沿。
       #执行定位 := #请求使能 AND NOT #执行标定 AND NOT #标定忙
       AND ((#状态 = 6) OR (#状态 = 21) OR (#状态 = 31));
       #执行停止 := #请求使能 AND NOT #执行标定 AND NOT #标定忙 AND (#状态 = 41);
       IF (#状态 = 6) OR (#状态 = 21) OR (#状态 = 31) THEN
           #动作计时 := "计时更新"(当前 := #动作计时, 步数 := #计时步数, 上限 := 12000);
           IF #动作计时 >= 12000 THEN
               #故障锁定 := TRUE;
               #故障码 := W#16#F003;
           END_IF;
       ELSE
           #动作计时 := 0;
       END_IF;
       IF #状态 = 41 THEN
           #停稳计时 := "计时更新"(当前 := #停稳计时, 步数 := #计时步数, 上限 := 1000);
           IF #停稳计时 >= 1000 THEN
               #故障锁定 := TRUE;
               #故障码 := W#16#F004;
           END_IF;
       ELSE
           #停稳计时 := 0;
       END_IF;

       // 【位移约束】每段目标是本次逻辑0～180范围，超过180+两倍容差的请求锁F008，提示坐标突变或起点异常。
       IF #执行定位 AND (ABS(#相对距离) > 180.0 + 2.0 * "右侧参数".到位允许误差) THEN
           #故障锁定 := TRUE;
           #故障码 := W#16#F008;
       END_IF;
       IF #故障锁定 THEN
           #状态 := 90;
           #启动完成 := FALSE;
           #请求使能 := FALSE;
           #执行定位 := FALSE;
           #执行停止 := FALSE;
       END_IF;

       // 【原生位置模式】车窗Power.StartMode=1，相对定位由MC_MoveRelative完成。
       "车窗使能"(Axis := "车窗轴",
              Enable := #请求使能,
              StartMode := 1,
              StopMode := 0,
              Status => #使能完成,
              Error => #使能出错,
              ErrorID => #使能错误码);
       "车窗复位"(Axis := "车窗轴",
              Execute := "右侧运行".复位请求,
              Restart := FALSE,
              Error => #复位出错,
              ErrorID => #复位错误码);
       #标定完成 := #执行标定;
       #标定忙 := FALSE;
       #标定出错 := FALSE;
       #标定错误码 := 0;
       "车窗相对定位"(Axis := "车窗轴",
                Execute := #执行定位,
                Distance := #相对距离,
                Velocity := #定位速度,
                Done => #定位完成,
                Busy => #定位忙,
                CommandAborted => #定位中断,
                Error => #定位出错,
                ErrorID => #定位错误码);
       "车窗停止"(Axis := "车窗轴",
              Execute := #执行停止,
              Done => #停止完成,
              Busy => #停止忙,
              Error => #停止出错,
              ErrorID => #停止错误码);

       IF #复位出错 THEN
           #故障锁定 := TRUE;
           #故障码 := #复位错误码;
       END_IF;
       IF #使能出错 AND (#复位等待计时 = 0) THEN
           #故障锁定 := TRUE;
           #故障码 := #使能错误码;
       END_IF;
       IF #定位出错 AND (#复位等待计时 = 0) THEN
           #故障锁定 := TRUE;
           #故障码 := #定位错误码;
       END_IF;
       IF #停止出错 AND (#复位等待计时 = 0) THEN
           #故障锁定 := TRUE;
           #故障码 := #停止错误码;
       END_IF;
       IF #标定出错 AND (#复位等待计时 = 0) THEN
           #故障锁定 := TRUE;
           #故障码 := #标定错误码;
       END_IF;

       IF #定位中断 AND ((#状态 = 6) OR (#状态 = 21) OR (#状态 = 31)) AND #请求使能 THEN
           #故障锁定 := TRUE;
           #故障码 := W#16#F006;
       END_IF;

       "右侧状态".车窗状态 := #状态;
       "右侧状态".车窗实际角度 := #角度;
       "右侧状态".车窗位置有效 := #反馈有效 AND #已有基准;
       "右侧状态".车窗启动完成 := #启动完成 AND NOT #故障锁定;
       "右侧状态".车窗故障码 := #故障码;
       // 【端点不能只靠四舍五入】0/100要求原生停稳和位置误差，运动中给1～99，反馈或启动无效时给255。
       #位置 := 255;
       IF "右侧状态".车窗位置有效 AND #启动完成 THEN
           IF #原生停稳 AND (ABS(#角度) <= "右侧参数".到位允许误差) THEN
               #位置 := 0;
           ELSIF #原生停稳 AND (ABS(#角度 - 180.0) <= "右侧参数".到位允许误差) THEN
               #位置 := 100;
           ELSE
               #开度整数 := REAL_TO_INT(#角度 / 180.0 * 100.0);
               IF #开度整数 < 1 THEN
                   #开度整数 := 1;
               END_IF;
               IF #开度整数 > 99 THEN
                   #开度整数 := 99;
               END_IF;
               #位置 := INT_TO_USINT(#开度整数);
           END_IF;
       END_IF;
       "右侧状态".车窗开度 := #位置;
END_FUNCTION_BLOCK

FUNCTION_BLOCK "右侧联动"   // FB3, SCL
{ S7_Optimized_Access := 'TRUE' }
VERSION : 5.0
// 文件定位：右PLC/10_右侧联动.scl；TIA块名：“右侧联动”。
//  本块属于V3简明；与另两版执行代码和参数完全相同，差别仅为注释组织。
//  建议从右PLC/00_Main.scl开始，再回到本块阅读。
   VAR_INPUT
      计时步数 : Int;
   END_VAR
   VAR
      接收帧 : Array[0..15] of Word;
      发送帧 : Array[0..15] of Word;
      曾经连接 : Bool;
      已见首帧 : Bool;
      上次心跳 : Word;
      心跳年龄 : Int := 30000;
      本机心跳 : Word;
      上次复位票号 : Word;
      通信停机锁定 : Bool;
      读结果 : Int;
      写结果 : Int;
   END_VAR
   VAR_TEMP
      帧有效 : Bool;
      新连接 : Bool;
      下标 : Int;
      位置 : USInt;
      数值 : Real;
   END_VAR
BEGIN
       // 职责：右PLC的通信入口和两个轴的唯一循环调度点。Main→右侧联动实例→雨刮器实例/车窗实例。
       // 本块先建立可信网络与控制条件，再执行两个FB，最后回传本扫描结果。命令和反馈各16个WORD即32字节。

       // 【本扫描先清脉冲】复位请求是一次事件，先清FALSE；只有新合法复位票出现且全释放时才在本扫描置TRUE。
       "右侧运行".复位请求 := FALSE;
       #心跳年龄 := "计时更新"(当前 := #心跳年龄, 步数 := #计时步数, 上限 := 30000);
       #读结果 := -1;
       IF "右侧参数".双机接收硬件标识 <> 0 THEN
           #读结果 := DPRD_DAT(LADDR := "右侧参数".双机接收硬件标识, RECORD => #接收帧);
       END_IF;
       #帧有效 := (#读结果 = 0) AND (#接收帧[0] = W#16#C401)
       AND (#接收帧[1] = W#16#0400) AND (#接收帧[2] = #接收帧[15])
       AND ((#接收帧[3] AND W#16#FFFC) = 0) AND (#接收帧[5] <= 1)
       AND (#接收帧[6] <= 3) AND (#接收帧[7] <= 1) AND (#接收帧[8] <= 1);
       FOR #下标 := 9 TO 14 DO
           IF #接收帧[#下标] <> 0 THEN
               #帧有效 := FALSE;
           END_IF;
       END_FOR;
       #新连接 := NOT #曾经连接 OR (#心跳年龄 >= 30);
       // 【首帧不启运动】首帧记心跳和复位票，后续变化心跳才确认通信。重连重建复位基线，不重放旧复位。
       IF #帧有效 THEN
           IF NOT #已见首帧 THEN
               #已见首帧 := TRUE;
               #上次心跳 := #接收帧[2];
               #上次复位票号 := #接收帧[4];
           ELSIF #接收帧[2] <> #上次心跳 THEN

               IF #新连接 THEN
                   #上次复位票号 := #接收帧[4];
               END_IF;
               #曾经连接 := TRUE;
               #心跳年龄 := 0;
               #上次心跳 := #接收帧[2];
           END_IF;
       END_IF;

       // 【通信看门狗】合法新心跳年龄<300 ms才在线；曾在线后失效锁存停机，网络恢复不自动清锁。
       "右侧运行".网络有效 := #曾经连接 AND (#心跳年龄 < 30) AND #帧有效;
       IF #曾经连接 AND NOT "右侧运行".网络有效 THEN
           #通信停机锁定 := TRUE;
       END_IF;

       // 【右侧复位核对】新复位票且运行许可、停止位、雨刷开关、车窗上下全为0，才解除通信锁并发MC复位事件。
       IF "右侧运行".网络有效 AND (#接收帧[4] <> #上次复位票号) THEN
           #上次复位票号 := #接收帧[4];
           IF NOT #接收帧[3].%X1 AND NOT #接收帧[3].%X0 AND (#接收帧[5] = 0)
               AND (#接收帧[7] = 0) AND (#接收帧[8] = 0) THEN
               #通信停机锁定 := FALSE;
               "右侧运行".复位请求 := TRUE;
           END_IF;
       END_IF;
       "右侧运行".联动许可 := "右侧运行".网络有效 AND #接收帧[3].%X0;
       "右侧运行".软件停止 := #通信停机锁定 OR #接收帧[3].%X1;
       "右侧运行".雨刷开关 := "右侧运行".网络有效 AND (#接收帧[5] = 1);
       "右侧运行".雨刷档位 := WORD_TO_INT(#接收帧[6]);
       "右侧运行".车窗向上 := "右侧运行".网络有效 AND (#接收帧[7] = 1);
       "右侧运行".车窗向下 := "右侧运行".网络有效 AND (#接收帧[8] = 1);

       // 【执行顺序】当前命令和许可已就绪；先雨刷，再车窗，两个FB都拿到本扫描同一时间步数。
       "雨刮器实例"(开关 := "右侧运行".雨刷开关,
               档位 := "右侧运行".雨刷档位,
               计时步数 := #计时步数);
       "车窗实例"(向上 := "右侧运行".车窗向上,
              向下 := "右侧运行".车窗向下,
              计时步数 := #计时步数,
              位置 => #位置);
       #本机心跳 := "字计数递增"(原值 := #本机心跳);
       FOR #下标 := 0 TO 15 DO
           #发送帧[#下标] := 0;
       END_FOR;
       // 【反馈先清再填】D401状态包含本扫描两个轴结果。字4开度255表示无效，字5完成次数只在整轮结束时变化。
       #发送帧[0] := W#16#D401;
       #发送帧[1] := W#16#0400;
       #发送帧[2] := #本机心跳;
       #发送帧[3] := #上次心跳;
       #发送帧[4] := 255;
       IF "右侧状态".车窗启动完成 AND "右侧状态".车窗位置有效 THEN
           #发送帧[4] := USINT_TO_WORD(#位置);
       END_IF;
       #发送帧[5] := "右侧状态".雨刷完成次数;
       #发送帧[6] := INT_TO_WORD("右侧状态".雨刷状态);
       #发送帧[7] := INT_TO_WORD("右侧状态".车窗状态);

       // 【角度封装】显示值×100转有符号INT再装进WORD；接收方先WORD_TO_INT再除100，不能按无符号解码负角度。
       IF "雨刮器实例".估算有效 THEN
           #数值 := LIMIT(MN := -327.68, IN := "雨刮器实例".估算角度, MX := 327.67);
           #发送帧[8] := INT_TO_WORD(REAL_TO_INT(#数值 * 100.0));
       END_IF;
       IF "右侧状态".车窗位置有效 THEN
           #数值 := LIMIT(MN := -327.68, IN := "右侧状态".车窗实际角度, MX := 327.67);
           #发送帧[9] := INT_TO_WORD(REAL_TO_INT(#数值 * 100.0));
       END_IF;

       // 【质量逐位解释】0雨刷实测有效（本版FALSE），1车窗实际反馈，2/3原生HomingDone，4/5各轴准备好，6通信锁，7雨刷估算。
       #发送帧[10].%X0 := FALSE;
       #发送帧[10].%X7 := "雨刮器实例".估算有效;
       #发送帧[10].%X1 := "右侧状态".车窗位置有效;
       #发送帧[10].%X2 := "雨刷轴".StatusBits.HomingDone;
       #发送帧[10].%X3 := "车窗轴".StatusBits.HomingDone;
       #发送帧[10].%X4 := "右侧状态".雨刷启动完成;
       #发送帧[10].%X5 := "右侧状态".车窗启动完成;
       #发送帧[10].%X6 := #通信停机锁定;
       #发送帧[11] := "右侧状态".雨刷故障码;
       #发送帧[12] := "右侧状态".车窗故障码;
       #发送帧[13] := DINT_TO_WORD("雨刷轴".StatusSensor[1].State);
       #发送帧[14] := DINT_TO_WORD("车窗轴".StatusSensor[1].State);
       #发送帧[15] := #本机心跳;
       #写结果 := -1;
       IF "右侧参数".双机发送硬件标识 <> 0 THEN
           #写结果 := DPWR_DAT(LADDR := "右侧参数".双机发送硬件标识, RECORD := #发送帧);
       END_IF;
END_FUNCTION_BLOCK

FUNCTION_BLOCK "扫描计时"   // FB4, SCL
{ S7_Optimized_Access := 'TRUE' }
VERSION : 5.0
// 文件定位：右PLC/01_扫描计时.scl；TIA块名：“扫描计时”。
//  本块属于V3简明；与另两版执行代码和参数完全相同，差别仅为注释组织。
//  建议从右PLC/00_Main.scl开始，再回到本块阅读。
   VAR_OUTPUT
      时间步数 : Int;
   END_VAR
   VAR
      时标 : LReal;
      不足十毫秒余量 : LReal;
      首次调用 : Bool := TRUE;
   END_VAR
   VAR_TEMP
      本周期秒 : LReal;
      完整步数 : DInt;
   END_VAR
BEGIN
       // 此FB把不固定的CPU扫描周期换算成统一10 ms步数。每个PLC都有自己的实例，不跨CPU共享时钟。
       // RUNTIME返回的是相邻调用之间的秒数，包含通信/中断消耗；首次只初始化，非正样本不累加。

       // 【计时来源】RUNTIME使用CPU时钟测相邻调用间隔，先读取再判断首样本；界面刷新快慢不会影响这里。
       #本周期秒 := RUNTIME(#时标);
       #时间步数 := 0;
       IF #首次调用 THEN
           #首次调用 := FALSE;
           #不足十毫秒余量 := 0.0;
       ELSIF #本周期秒 > 0.0 THEN
           #不足十毫秒余量 := #不足十毫秒余量 + #本周期秒;

           // 【饱和】300 s相当于30000个10 ms步，仍在INT正范围内，防止暂停后转换溢出。
           IF #不足十毫秒余量 >= 300.0 THEN
               #时间步数 := 30000;
               #不足十毫秒余量 := 0.0;
           ELSE
               // 【保留余量】只输出完整10 ms的部分，减去已输出时间，未满一格的余量下次继续用。
               #完整步数 := TRUNC_DINT(#不足十毫秒余量 / 0.01);
               #时间步数 := DINT_TO_INT(#完整步数);
               #不足十毫秒余量 := #不足十毫秒余量 - DINT_TO_LREAL(#完整步数) * 0.01;
           END_IF;
       END_IF;
END_FUNCTION_BLOCK

FUNCTION "字计数递增" : Word   // FC1, SCL
{ S7_Optimized_Access := 'TRUE' }
VERSION : 4.0
// 汽车综合实践完整中文版 V4.0；所有自定义名称与注释使用中文。
//  导入前：先建立“雨刷轴”“车窗轴”两个软件工艺对象；再按指南创建九个运动指令实例。
//  报文3由工艺对象独占。严禁另行写入驱动输出字；本文件无外接传感器地址。
   VAR_INPUT
      原值 : Word;
   END_VAR
BEGIN
       IF #原值 = W#16#FFFF THEN
           #字计数递增 := 0;
       ELSE
           #字计数递增 := UINT_TO_WORD(WORD_TO_UINT(#原值) + UINT#1);
       END_IF;
END_FUNCTION

FUNCTION "计时更新" : Int   // FC2, SCL
{ S7_Optimized_Access := 'TRUE' }
VERSION : 5.0
// 文件定位：右PLC/03_计时更新.scl；TIA块名：“计时更新”。
//  本块属于V3简明；与另两版执行代码和参数完全相同，差别仅为注释组织。
//  建议从右PLC/00_Main.scl开始，再回到本块阅读。
   VAR_INPUT
      当前 : Int;
      步数 : Int;
      上限 : Int;
   END_VAR
   VAR_TEMP
      新值 : DInt;
   END_VAR
BEGIN
       // 公共饱和计时FC，没有独立历史记忆：输入当前值、增量和上限，返回0～上限的INT。
       // 先把两个INT转DINT相加，再LIMIT，最后转回INT；加法不会先在INT中溢出。

       #新值 := INT_TO_DINT(#当前) + INT_TO_DINT(#步数);
       #计时更新 := DINT_TO_INT(LIMIT(MN := DINT#0, IN := #新值, MX := INT_TO_DINT(#上限)));
END_FUNCTION

ORGANIZATION_BLOCK "Main"   // OB1, SCL, ProgramCycle
{ S7_Optimized_Access := 'TRUE' }
VERSION : 5.0
// 文件定位：右PLC/00_Main.scl；TIA块名：“Main”。
//  本块属于V3简明；与另两版执行代码和参数完全相同，差别仅为注释组织。
   VAR_INPUT
      Initial_Call : Bool;   // Initial call of this OB
      Remanence : Bool;   // =True, if remanent data are available
   END_VAR
   VAR_TEMP
      时间步数 : Int;
   END_VAR
BEGIN
       // 阅读入口：本文件是右PLC的Main循环组织块。完整源在“右PLC_完整.scl”，分块入口在“右PLC/00_Main.scl”。
       // 调用顺序：Main → 扫描计时实例（FB扫描计时）→ 右侧联动实例（FB右侧联动）。
       // Main每扫描只获取一次时间，然后把同一时间步数传给本PLC的全部业务。时间步数为0也照常调用业务。
       // 第一跳：右PLC/01_扫描计时.scl；第二跳：右PLC/10_右侧联动.scl；第三跳：右PLC/03_计时更新.scl。
       // 实例DB说明分别在右PLC/02_扫描计时实例.scl、右PLC/11_右侧联动实例.scl。
       // 雨刷每半程小15 s、中10 s、大5 s；一次固定中档，正反向命令共20 s，换向仍等待原生停稳。
       // 车窗使用实际反馈的相对坐标，默认45度/秒，方向系数同时作用于指令与反馈。
       // 默认无手操盒。先释放动作与控制申请，复位得到接受后再申请运行。

       "扫描计时实例"(时间步数 => #时间步数);

       "右侧联动实例"(计时步数 := #时间步数);
END_ORGANIZATION_BLOCK

ORGANIZATION_BLOCK "启动初始化"   // OB100, SCL, Startup
{ S7_Optimized_Access := 'TRUE' }
VERSION : 5.0
// 文件定位：右PLC/90_启动初始化.scl；TIA块名：“启动初始化”。
//  本块属于V3简明；与另两版执行代码和参数完全相同，差别仅为注释组织。
//  建议从右PLC/00_Main.scl开始，再回到本块阅读。
   VAR_INPUT
      LostRetentive : Bool;   // True if retentive data are lost
      LostRTC : Bool;   // True if date and time are lost
   END_VAR
BEGIN
       // CPU启动时清通信基线、动作和时基，先锁停；复位接受后再申请控制。

       "右侧参数".实机调试完成 := FALSE;
       "右侧参数".维护模式 := FALSE;
       "右侧参数".雨刷标定申请 := FALSE;
       "右侧参数".车窗标定申请 := FALSE;
       "右侧运行".联动许可 := FALSE;
       "右侧运行".复位请求 := FALSE;
       "右侧运行".软件停止 := TRUE;
       "右侧运行".网络有效 := FALSE;
       "右侧联动实例".曾经连接 := FALSE;
       "右侧联动实例".已见首帧 := FALSE;
       "右侧联动实例".心跳年龄 := 30000;

       "右侧联动实例".通信停机锁定 := TRUE;
       "雨刮器实例".状态 := 0;
       "雨刮器实例".相对基准有效 := FALSE;
       "雨刮器实例".估算有效 := FALSE;
       "雨刮器实例".上次标定申请 := FALSE;
       "雨刮器实例".启动完成 := FALSE;
       "车窗实例".状态 := 0;
       "车窗实例".相对基准有效 := FALSE;
       "车窗实例".上次标定申请 := FALSE;
       "车窗实例".启动完成 := FALSE;
       "右侧状态".雨刷位置有效 := FALSE;
       "右侧状态".车窗位置有效 := FALSE;
       "右侧状态".雨刷启动完成 := FALSE;
       "右侧状态".车窗启动完成 := FALSE;
       "右侧状态".车窗开度 := 255;

       "扫描计时实例".时标 := 0.0;
       "扫描计时实例".不足十毫秒余量 := 0.0;
       "扫描计时实例".首次调用 := TRUE;
       "扫描计时实例".时间步数 := 0;
END_ORGANIZATION_BLOCK

(* ===== HMI "HMI_RT_1" =====
system functions are stored by id; their names below are inferred from use
connection "连接_PLC左_集成": ETHERNET, SMART_S7_1200_OMS

HMI tags "默认变量表"
   "Tag_ScreenNumber" : UInt, internal

HMI tags "汽车控制变量"
   "有效雨刷模式" : UInt AT %DB101.DBW14, 100 ms   // 只读；DB101.DBW14
   "有效雨刷档位" : UInt AT %DB101.DBW16, 100 ms   // 只读；DB101.DBW16
   "车窗状态" : UInt AT %DB101.DBW68, 100 ms   // 只读；DB101.DBW68
   "允许面板操作" : Bool AT %DB101.DBX39.0, 100 ms   // 只读；DB101.DBX39.0
   "允许一次雨刷" : Bool AT %DB101.DBX39.1, 100 ms   // 只读；DB101.DBX39.1
   "允许面板升降" : Bool AT %DB101.DBX39.2, 100 ms   // 只读；DB101.DBX39.2
   "两轴启动完成" : Bool AT %DB101.DBX25.6, 100 ms   // 只读；DB101.DBX25.6
   "雨刷故障码" : UInt AT %DB101.DBW70, 100 ms   // 只读；DB101.DBW70
   "车窗故障码" : UInt AT %DB101.DBW72, 100 ms   // 只读；DB101.DBW72
   "关挡票" : Bool AT %DB102.DBX1.0, 100 ms   // 面板独占写；DB102.DBX1.0
   "自动票" : Bool AT %DB102.DBX3.0, 100 ms   // 面板独占写；DB102.DBX3.0
   "小挡票" : Bool AT %DB102.DBX5.0, 100 ms   // 面板独占写；DB102.DBX5.0
   "中挡票" : Bool AT %DB102.DBX7.0, 100 ms   // 面板独占写；DB102.DBX7.0
   "大挡票" : Bool AT %DB102.DBX9.0, 100 ms   // 面板独占写；DB102.DBX9.0
   "一次票" : Bool AT %DB102.DBX11.0, 100 ms   // 面板独占写；DB102.DBX11.0
   "面板向上保持" : Bool AT %DB102.DBX13.0, 100 ms   // 面板独占写；DB102.DBX13.0
   "面板向下保持" : Bool AT %DB102.DBX15.0, 100 ms   // 面板独占写；DB102.DBX15.0
   "面板控制会话请求" : Bool AT %DB102.DBX23.0, 100 ms   // 面板独占写；DB102.DBX23.0
   "复位票" : Bool AT %DB102.DBX19.0, 100 ms   // 面板独占写；DB102.DBX19.0
   "软件停止票" : Bool AT %DB102.DBX21.0, 100 ms   // 面板独占写；DB102.DBX21.0
   "面板当前画面" : UInt AT %DB102.DBW26, 100 ms   // 面板独占写；DB102.DBW26
   "雨刷就绪" : Bool AT %DB101.DBX79.2, 100 ms   // 只读；DB101.DBX79.2；字[39]独立轴就绪反馈
   "车窗就绪" : Bool AT %DB101.DBX79.3, 100 ms   // 只读；DB101.DBX79.3；字[39]独立轴就绪反馈
   "车窗当前角度" : Int AT %DB101.DBW60, 100 ms   // 只读车窗反馈；%DB101.DBW60
   "车窗当前开度" : UInt AT %DB101.DBW32, 100 ms   // 只读车窗反馈；%DB101.DBW32
   "车窗位置有效" : Bool AT %DB101.DBX63.1, 100 ms   // 只读车窗反馈；%DB101.DBX63.1

text list "单页_雨刷模式": 0 '关'; 1 '自动'; 2 '小'; 3 '中'; 4 '大'

text list "单页_雨刷档位": 0 '停止'; 1 '低档'; 2 '中档'; 3 '高档'

text list "单页_车窗状态": 0 '未就绪'; 5 '回位'; 6 '回位'; 10 '停止'; 20 '上行'; 21 '上行'; 30 '下行'; 31 '下行'; 40 '停止中'; 41 '停止中'; 90 '故障'

text list "单页_控制许可": 0 '未获控制'; 1 '已获控制'

text list "单页_系统就绪": 0 '雨刷/车窗未就绪'; 1 '雨刷/车窗已就绪'

text list "单页_雨刷就绪": 0 '雨刷未就绪'; 1 '雨刷已就绪'

text list "单页_车窗就绪": 0 '车窗未就绪'; 1 '车窗已就绪'

Template "模板_1" 800x480
   Button "退出" at 714,429 size 71x50; TextOff '退出'; PictureOff "ExitRuntime_KTP700_Basic_PN_TR"; PictureOn "ExitRuntime_KTP700_Basic_PN_TR"
      on Release: StopRuntime(0)
   Button "Template_Button" at 614,429 size 71x50; TextOff 'Text'
   Button "Template_Button_1" at 514,429 size 71x50; TextOff 'Text'
   Button "Template_Button_2" at 414,429 size 71x50; TextOff 'Text'
   Button "Template_Button_3" at 314,429 size 71x50; TextOff 'Text'
   Button "Template_Button_4" at 214,429 size 71x50; TextOff 'Text'
   Button "报警" at 114,429 size 71x50; TextOff '报警'; PictureOff "AlarmDisplay_KTP700_Basic_PN_TR"; PictureOn "AlarmDisplay_KTP700_Basic_PN_TR"
      on Release: function_ef3f5d25("报警窗口_Unacknowledged", -1)
   Button "起始画面" at 14,429 size 71x50; TextOff '起始画面'; PictureOff "NavigateHome_KTP700_Basic_PN_TR"; PictureOn "NavigateHome_KTP700_Basic_PN_TR"
      on Release: ActivateScreen("根画面", 0)
   SymbolicIOField "Symbolic_IO_Field_Screen" at 93,9 size 600x33; TextOff '0'; TextOn '1'; TextList "TextList_ScreenNames"
      ProcessValue <- "Tag_ScreenNumber"
      on Change: ActivateScreenByNumber("Tag_ScreenNumber", 0)
   DateTimeField "HmiScreenItemData" at 695,25 size 105x25
   DateTimeField "HmiScreenItemData_1" at 695,0 size 105x25
   GraphicView "Logo" at 0,0 size 91x51; Picture "HMI_1 的 Logo"

screen "根画面" 800x480
   on ClearScreen: ResetBit("面板向上保持"); ResetBit("面板向下保持")
   on GenerateScreen: SetTag("面板当前画面", 0); ResetBit("面板向上保持"); ResetBit("面板向下保持")
   TextField "标题" at 24,16 size 300x36; Text '汽车控制'
   SymbolicIOField "控制权限" at 558,18 size 218x34; TextOff '0'; TextOn '1'; TextList "单页_控制许可"
      ProcessValue <- "允许面板操作"
   TextField "雨刷分组" at 24,78 size 74x28; Text '雨刷'
   TextField "模式标签" at 110,80 size 48x26; Text '模式'
   SymbolicIOField "最终雨刷模式" at 164,76 size 116x34; TextOff '0'; TextOn '1'; TextList "单页_雨刷模式"
      ProcessValue <- "有效雨刷模式"
   TextField "档位标签" at 300,80 size 48x26; Text '档位'
   SymbolicIOField "最终雨刷档位" at 354,76 size 138x34; TextOff '0'; TextOn '1'; TextList "单页_雨刷档位"
      ProcessValue <- "有效雨刷档位"
   TextField "车窗分组" at 532,78 size 70x28; Text '车窗'
   SymbolicIOField "最终车窗状态" at 610,76 size 166x34; TextOff '0'; TextOn '1'; TextList "单页_车窗状态"
      ProcessValue <- "车窗状态"
   Button "雨刷关" at 24,130 size 148x72; TextOff '关'
      on Click: InvertBit("关挡票")
   Button "雨刷自动" at 184,130 size 148x72; TextOff '自动'
      on Click: InvertBit("自动票")
   Button "雨刷小" at 24,218 size 148x72; TextOff '小'
      on Click: InvertBit("小挡票")
   Button "雨刷中" at 184,218 size 148x72; TextOff '中'
      on Click: InvertBit("中挡票")
   Button "雨刷大" at 344,218 size 148x72; TextOff '大'
      on Click: InvertBit("大挡票")
   Button "雨刷一次" at 344,130 size 148x72; TextOff '一次'
      on Click: InvertBit("一次票")
   Button "车窗上行" at 532,130 size 244x72; TextOff '上行'
      on Press: SetBit("面板向上保持")
      on Release: ResetBit("面板向上保持")
   Button "车窗下行" at 532,218 size 244x72; TextOff '下行'
      on Press: SetBit("面板向下保持")
      on Release: ResetBit("面板向下保持")
   SymbolicIOField "雨刷就绪" at 24,326 size 228x36; TextOff '0'; TextOn '1'; TextList "单页_雨刷就绪"
      ProcessValue <- "雨刷就绪"
   SymbolicIOField "车窗就绪" at 532,326 size 244x36; TextOff '0'; TextOn '1'; TextList "单页_车窗就绪"
      ProcessValue <- "车窗就绪"
   TextField "雨刷故障提示" at 24,362 size 228x24; Text '雨刷故障'
      Visibility <- "雨刷故障码"
   TextField "车窗故障提示" at 532,362 size 244x24; Text '车窗故障'
      Visibility <- "车窗故障码"
   Button "复位" at 344,390 size 156x66; TextOff '复位'
      on Click: ResetBit("面板控制会话请求"); ResetBit("面板向上保持"); ResetBit("面板向下保持"); InvertBit("复位票")
   Button "软件停止" at 520,390 size 256x66; TextOff '软件停止'
      on Click: ResetBit("面板控制会话请求"); ResetBit("面板向上保持"); ResetBit("面板向下保持"); InvertBit("软件停止票")
   TextField "车窗位置标签" at 532,296 size 46x28; Text '位置'
   IOField "车窗角度值" at 580,296 size 84x28; FormatPattern 999
      ProcessValue <- "车窗当前角度"
      Visibility <- "车窗位置有效"
   IOField "车窗开度值" at 690,296 size 58x28; FormatPattern 999
      ProcessValue <- "车窗当前开度"
      Visibility <- "车窗位置有效"
   TextField "车窗角度单位" at 666,296 size 18x28; Text '°'
      Visibility <- "车窗位置有效"
   TextField "车窗开度单位" at 751,296 size 23x28; Text '%'
      Visibility <- "车窗位置有效"
   TextField "车窗位置无效提示" at 580,296 size 194x28; Text '位置未就绪'
      Visibility <- "车窗位置有效"
   Button "申请控制按钮" at 24,390 size 300x66; TextOff '申请控制'
      on Click: InvertBit("面板控制会话请求")
      Visibility <- "面板控制会话请求"
   Button "释放控制按钮" at 24,390 size 300x66; TextOff '释放控制'
      on Click: InvertBit("面板控制会话请求")
      Visibility <- "面板控制会话请求"
*)